(* IEC 61131-3 sources: JingjiangArm/moonboxpro_arm_8.4/Application/Application/任务列表/TensionTask/张力控制/收放料/张力调整/Tension_2024, 5 files *)

(* ---- KS_InitTensionCtl_StructParam.st ---- *)
(*@CES
Name=KS_InitTensionCtl_StructParam
Type=FunctionBlock
TypeGuid=6f9dac99-8de1-4efc-8465-68ac443b7d08
Guid=d3edacb8-afe0-4e68-804f-3598657c3108
HasDeclaration=True
HasImplementation=True
*)
{DECLARATION}
FUNCTION KS_InitTensionCtl_StructParam : BOOL(*初始化张力控制结构体参数*)
VAR_INPUT
	i_byInitEn:BYTE;(*初始化使能标志@按照定义顺序/.0 初始化第一个结构体。以此类推！*)
	i_xUseIMatrix_rX_DARE:BOOL;(*迭代计算的初始矩阵为单位矩阵@否则为特定初始卷径的收敛值*)
	(*/.0*)
	i_pstInitial_Model_Parameters_Input: POINTER TO Initial_Model_Parameters;(*2024.05.07.093000 调整接口名*)
	(*/.1*)
	i_pstInvariant_Parameters1: POINTER TO Invariant_Parameters;(*2024.05.07.105319 修改接口名by Liu*)
	(*/.2*)
	i_pstKalman_Status_Estimation_And_Feedback1: POINTER TO Kalman_Status_Estimation_And_Feedback;(*2024.05.07.105319 修改接口名by Liu*)
	(*/.3*)
	i_pstKalman_Status_Estimation_And_Feedback_MinBeat1: POINTER TO Kalman_Status_Estimation_And_Feedback_MinBeat;(*2024.05.07.105319 修改接口名by Liu*)
	(*/.4*)
	i_pstPI_Parameters1: POINTER TO PI_Parameters;(*2024.05.07.105319 修改接口名by Liu*)
	(*LQR迭代求解DARE@函数中初始化为了特定初始卷径的收敛值|
	如果初始化为了单位矩阵，需要迭代，第一拍迭代可能时间会长*)
	(*2024.06.08.151322 修改为了lreal类型*)
	(*/.5*)
	i_parX_DARE:POINTER TO ARRAY [1..4,1..4] OF REAL;(*上一个周期已经迭代收敛的值X_Dare*)
	i_palrX_DARE:POINTER TO ARRAY [1..4,1..4] OF LREAL;(*上一个周期已经迭代收敛的值X_Dare*)
	(*/.6@2024.05.13.181113+*)
	i_pstPI_Parameters1_AccDec: POINTER TO PI_Parameters;(*2024.05.13.181126 升降速pi参数*)
	i_iCycleTime_Plc: INT;
END_VAR
VAR
	xInit: BOOL;
	arQ:ARRAY [1..4,1..4] OF REAL;(*Q矩阵*)
	arI:ARRAY [1..4,1..4] OF REAL;(*单位矩阵*)
	arKf:ARRAY [1..4] OF REAL;
	arX_DARE:ARRAY [1..4,1..4] OF REAL;
	(*2024.06.08.151416增加lreal类型*)
	alrQ:ARRAY [1..4,1..4] OF LREAL;(*Q矩阵*)
	alrKf:ARRAY [1..4] OF LREAL;
	alrI:ARRAY [1..4,1..4] OF LREAL;(*单位矩阵*)
	alrX_DARE:ARRAY [1..4,1..4] OF LREAL;
END_VAR
{IMPLEMENTATION}
(*初始化第一个结构体*)
xInit:=i_byInitEn.0;
IF i_pstInitial_Model_Parameters_Input<>0 AND xInit THEN
   	i_pstInitial_Model_Parameters_Input^.R_0	:=0.27;             (*初始卷半径m 0.31*)

    i_pstInitial_Model_Parameters_Input^.a0_0	:=0;           	(*初始a0*)
    i_pstInitial_Model_Parameters_Input^.b1_0	:=0.07;	 			(*初始b1 0.016*)
    i_pstInitial_Model_Parameters_Input^.Wn_0	:=8.9;				(*初始Wn 4.3*)
    i_pstInitial_Model_Parameters_Input^.Beta_0	:=0.5;				(*初始Beta  0.22*)

    i_pstInitial_Model_Parameters_Input^.l_0	:=1;				(*初始调整系数l 1*)
END_IF

(*初始化第二个结构体*)
xInit:=i_byInitEn.1;
IF i_pstInvariant_Parameters1<>0 AND xInit THEN
    i_pstInvariant_Parameters1^.Ts		:=INT_TO_REAL(i_iCycleTime_Plc)/1000.0;		(*采样时间Ts*)
    i_pstInvariant_Parameters1^.Range	:=11.8;    	(*输出最大量程 13.8*)
    i_pstInvariant_Parameters1^.Theta	:=30.0;	(*摆臂偏角范围 25.64*)

    i_pstInvariant_Parameters1^.K_adj	:=1.4;		(*模型调整增益 1.3*)
END_IF

(*构造一个单位矩阵*)
arI[1,1]:=1;
arI[2,2]:=1;
arI[3,3]:=1;
arI[4,4]:=1;
alrI[1,1]:=1;
alrI[2,2]:=1;
alrI[3,3]:=1;
alrI[4,4]:=1;
(*构造一个Q矩阵*)
arQ[4,4]:=0.01;
alrQ[4,4]:=0.01;
(*构造kf矩阵*)
arKf[1]:=-0.71625816;
arKf[2]:=-14.455574;
arKf[3]:=-25.065932;
arKf[4]:=-341.98005;

alrKf[1]:=-0.71625816;
alrKf[2]:=-14.455574;
alrKf[3]:=-25.065932;
alrKf[4]:=-341.98005;

(*初始化第三个结构体*)
xInit:=i_byInitEn.2;
IF i_pstKalman_Status_Estimation_And_Feedback1<>0 AND xInit THEN
	i_pstKalman_Status_Estimation_And_Feedback1^.R_K	:=10;
	i_pstKalman_Status_Estimation_And_Feedback1^.Q		:=arQ;
	i_pstKalman_Status_Estimation_And_Feedback1^.P0		:=arI;
	i_pstKalman_Status_Estimation_And_Feedback1^.N_LQR	:=10;
	i_pstKalman_Status_Estimation_And_Feedback1^.Kf		:=arKf;

	i_pstKalman_Status_Estimation_And_Feedback1^.alrQ		:=alrQ;
	i_pstKalman_Status_Estimation_And_Feedback1^.alrP0		:=alrI;
	i_pstKalman_Status_Estimation_And_Feedback1^.alrKf		:=alrKf;
END_IF

(*初始化第四个结构体*)
xInit:=i_byInitEn.3;
IF i_pstKalman_Status_Estimation_And_Feedback_MinBeat1<>0 AND xInit THEN
	i_pstKalman_Status_Estimation_And_Feedback_MinBeat1^.R_K	:=100;
	i_pstKalman_Status_Estimation_And_Feedback_MinBeat1^.Q		:=arQ;
	i_pstKalman_Status_Estimation_And_Feedback_MinBeat1^.P0		:=arI;
	i_pstKalman_Status_Estimation_And_Feedback_MinBeat1^.N_MinBeat:=2;
	i_pstKalman_Status_Estimation_And_Feedback_MinBeat1^.Kf		:=arKf;
END_IF

(*初始化第五个结构体*)
xInit:=i_byInitEn.4;
IF i_pstPI_Parameters1<>0 AND xInit THEN
	i_pstPI_Parameters1^.K_PI	:=1;
	i_pstPI_Parameters1^.a		:=4.2;

	i_pstPI_Parameters1^.b		:=0;
END_IF

(*初始化第六个结构体*)
(*构造arX_DARE矩阵@特定初始卷径的收敛值*)

arX_DARE[1,1]:=0.5809964918;
arX_DARE[1,2]:=11.4605492993;
arX_DARE[1,3]:=19.3883120752;
arX_DARE[1,4]:=261.7670536474;

arX_DARE[2,1]:=11.4605492993;
arX_DARE[2,2]:=341.4559372966;
arX_DARE[2,3]:=273.7038620995;
arX_DARE[2,4]:=2799.1520439073;

arX_DARE[3,1]:=19.3883120752;
arX_DARE[3,2]:=273.7038620995;
arX_DARE[3,3]:=758.807264184;
arX_DARE[3,4]:=11796.8531367233;

arX_DARE[4,1]:=261.7670536474;
arX_DARE[4,2]:=2799.1520439073;
arX_DARE[4,3]:=11796.8531367233;
arX_DARE[4,4]:=347613.458626343;

(*LREAL*)
alrX_DARE[1,1]:=0.5809964918;
alrX_DARE[1,2]:=11.4605492993;
alrX_DARE[1,3]:=19.3883120752;
alrX_DARE[1,4]:=261.7670536474;

alrX_DARE[2,1]:=11.4605492993;
alrX_DARE[2,2]:=341.4559372966;
alrX_DARE[2,3]:=273.7038620995;
alrX_DARE[2,4]:=2799.1520439073;

alrX_DARE[3,1]:=19.3883120752;
alrX_DARE[3,2]:=273.7038620995;
alrX_DARE[3,3]:=758.807264184;
alrX_DARE[3,4]:=11796.8531367233;

alrX_DARE[4,1]:=261.7670536474;
alrX_DARE[4,2]:=2799.1520439073;
alrX_DARE[4,3]:=11796.8531367233;
alrX_DARE[4,4]:=347613.458626343;

xInit:=i_byInitEn.5;
IF i_parX_DARE<>0 AND xInit THEN
	IF i_xUseIMatrix_rX_DARE THEN(*初始化单位矩阵*)
		i_parX_DARE^:=arI;
	ELSE(*初始化为特定初始卷径的收敛值*)
		i_parX_DARE^:=arX_DARE;
	END_IF
END_IF
IF i_palrX_DARE<>0 AND xInit THEN
	IF i_xUseIMatrix_rX_DARE THEN(*初始化单位矩阵*)
		i_palrX_DARE^:=alrI;
	ELSE(*初始化为特定初始卷径的收敛值*)
		i_palrX_DARE^:=alrX_DARE;
	END_IF
END_IF

(*初始化第七个结构体*)
xInit:=i_byInitEn.6;
IF i_pstPI_Parameters1_AccDec<>0 AND xInit THEN
	i_pstPI_Parameters1_AccDec^.K_PI	:=1;
	i_pstPI_Parameters1_AccDec^.a		:=7.2;
	i_pstPI_Parameters1_AccDec^.b		:=0;
END_IF

(* ---- Para_Cal.st ---- *)
(*@CES
Name=Para_Cal
Type=FunctionBlock
TypeGuid=6f9dac99-8de1-4efc-8465-68ac443b7d08
Guid=ef90c73f-dc4b-4bec-847d-13655df4417f
HasDeclaration=True
HasImplementation=True
*)
{DECLARATION}
FUNCTION Para_Cal : REAL
(*做了微调@2024.05.07.103831by Liu*)
(*主要是用于使用时变参数/设置参数的切换*)
(*时变算法还不太完善，需要优化切记！！！@2024.05.13.193242*)
(*2025.5.12.211538 限制不能为负值*)
VAR_INPUT
	i_xUseTime_Variaition:BOOL;(*使用时变算法*)
	i_stInitial_Model_Parameters_Input: Initial_Model_Parameters;(*2024.05.07.093000 调整接口名*)
	i_pTime_Varying_Parameters_Output: POINTER TO Time_Varying_Parameters;
	i_rEST_R:REAL;(*估计的卷半径m*)
	i_rUseTime_R_Min:REAL;(*使用时变的最小卷半径|m@2024.05.14.080937*)
	i_xUseTime_b1:BOOL;(*有效则b1随卷径实时变化-不实时变化则使用b1_0@2024.05.14.080937*)
END_VAR

VAR
	(*2024.05.07.092928 调整@Liu*)
	Initial_Model_Parameters_Input: Initial_Model_Parameters;
	rE:REAL:=2.718281828459045;(*自然常数e*)
(*Initial_Model_Parameters*)
	R_0: REAL;             (*初始卷半径m*)
	a0_0: REAL;           (*初始a0*)
	b1_0: REAL;	 	(*初始b1*)
	Wn_0: REAL;	(*初始Wn*)
	Beta_0: REAL;	(*初始Beta*)
	l_0: REAL;		(*初始调整系数l*)
(*Time_Varying_Parameters*)
	Ru:REAL;(*估计的卷半径m*)
	a0:REAL;
	b1:REAL;
	Beta:REAL;
	Wn:REAL;
	l:REAL;
(*中间变量*)
	Temp:REAL;
	Ru_Temp:REAL;
	rUseTime_R_Min: REAL;
END_VAR
{IMPLEMENTATION}
	rUseTime_R_Min:=i_rUseTime_R_Min;
	IF rUseTime_R_Min<95.0/2/1000 THEN(*做合法判断*)
		rUseTime_R_Min:=95.0/2/1000;
	END_IF

	(*内部参数赋值*)
	Initial_Model_Parameters_Input:=i_stInitial_Model_Parameters_Input;(*2024.05.07.092953|liu*)
	(*Initial_Model_Parameters*)
	R_0  	:= Initial_Model_Parameters_Input.R_0;             (*初始卷半径m*)
	IF R_0<90.0/2/1000 THEN(*初始卷径默认值@2024.05.07.103750|下面逻辑有/的操作*)
		R_0:=90.0/2/1000;
	END_IF

	a0_0	:= Initial_Model_Parameters_Input.a0_0;           (*初始a0*)
	b1_0 	:= Initial_Model_Parameters_Input.b1_0;	 	(*初始b1*)
	Wn_0 	:= Initial_Model_Parameters_Input.Wn_0;	(*初始Wn*)
	Beta_0 	:= Initial_Model_Parameters_Input.Beta_0;	(*初始Beta*)
	l_0 	:= Initial_Model_Parameters_Input.l_0;		(*初始调整系数l*)
	(*半径*)
	(*Ru 计算主机转速@重要*)
	Ru := i_rEST_R;

	IF i_xUseTime_Variaition THEN(*使用估计的转速值到电机*);
		(*根据卷径关系计算时变参数*)
(*
	(*	b1 := b1_0*EXPT((R_0/Ru),3); *)
		Temp := -3.99*(Ru/R_0);
(*		b1 := 0.8648 * EXPT(gc_rE,Temp);*)
(*		b1 := 0.8648 * EXPT(rE,Temp);*)
		b1 :=0.05;(*华丰测试使用@2024.05.13.193222*)
		Beta := Beta_0*EXPT((R_0/Ru),2);
		Wn := Wn_0*EXPT((R_0/Ru),2);
		l := l_0;
		a0 := a0_0;
*)

		(*根据卷径关系计算时变参数  考虑小卷时转动惯量不随Ru变化 对Ru做判断*)
		(*Ru_Temp 用于计算时变参数*)
		IF Ru<rUseTime_R_Min THEN(*初始卷径默认值@2024.05.07.103750|下面逻辑有/的操作*)
			Ru_Temp:=rUseTime_R_Min;
		ELSE
			Ru_Temp:=Ru;
		END_IF

	(*	b1 := b1_0*EXPT((R_0/Ru),3); *)
		Temp := -3.99*(Ru_Temp/R_0);
		IF i_xUseTime_b1 THEN
			b1 := 0.8648 * EXPT(rE,Temp);
			(*2025.5.12.211538 限制不能为负值*)
			IF b1<=0 THEN
				b1:=0.01;
			END_IF
		ELSE
			b1 :=b1_0;(*华丰测试使用@2024.05.13.193222*)
		END_IF
		Beta := LREAL_TO_REAL(Beta_0*EXPT((R_0/Ru_Temp),2));
		Wn := LREAL_TO_REAL(Wn_0*EXPT((R_0/Ru_Temp),2));
		l := l_0;
		a0 := a0_0;

		(*结构体赋值*)
		i_pTime_Varying_Parameters_Output^.EST_R := Ru;
		i_pTime_Varying_Parameters_Output^.a0 := a0;
		i_pTime_Varying_Parameters_Output^.b1 := b1;
		i_pTime_Varying_Parameters_Output^.Wn := Wn;
		i_pTime_Varying_Parameters_Output^.Beta := Beta;
		i_pTime_Varying_Parameters_Output^.l := l;
	ELSE
		(*结构体赋值*)
		i_pTime_Varying_Parameters_Output^.EST_R := Ru;
		i_pTime_Varying_Parameters_Output^.a0 := a0_0;
		i_pTime_Varying_Parameters_Output^.b1 := b1_0;
		i_pTime_Varying_Parameters_Output^.Wn := Wn_0;
		i_pTime_Varying_Parameters_Output^.Beta := Beta_0;
		i_pTime_Varying_Parameters_Output^.l := l_0;
	END_IF

(* ---- Time_Variaition_PILQR.st ---- *)
(*@CES
Name=Time_Variaition_PILQR
Type=FunctionBlock
TypeGuid=6f9dac99-8de1-4efc-8465-68ac443b7d08
Guid=72ca66b0-1667-4547-85f7-d4b61b3bde5a
HasDeclaration=True
HasImplementation=True
*)
{DECLARATION}
FUNCTION Time_Variaition_PILQR : REAL
VAR_INPUT
	i_xUseWfValue:BOOL;(*使用估计的转速值到电机|不使用的时候清除估计转速输出*)
(*输入变量*)
	i_rVt:REAL;(*牵引线速度m/min*)
	i_rWu:REAL;(*放料转速(RPM)*)
	i_rY:REAL;(*张力摆臂反馈*)
	i_rKc: REAL;		(*调整增益*)
(*输出变量指针*)
	i_piK:POINTER TO INT;(*拍数计数*)
	i_prWf:POINTER TO REAL;(*转速补偿量r/min*)
	i_prCNT:POINTER TO REAL;(*LQR迭代次数*)
(*结构体*)
	i_stInvariant_Parameters1:Invariant_Parameters;(*2024.05.07.105319 修改接口名by Liu*)
	i_stTime_Varying_Parameters1:Time_Varying_Parameters;(*2024.05.07.105319 修改接口名by Liu*)
	i_stKalman_Status_Estimation_And_Feedback1:Kalman_Status_Estimation_And_Feedback;(*2024.05.07.105319 修改接口名by Liu*)
	i_stPI_Parameters1:PI_Parameters;(*2024.05.07.105319 修改接口名by Liu*)
	i_pCached_Array_Pointers1: POINTER TO Cached_Array_Pointers;
END_VAR

VAR
	(*2024.05.07.105252 增加局部变量by Liu*)
	Invariant_Parameters1:Invariant_Parameters;
	Time_Varying_Parameters1:Time_Varying_Parameters;
	Kalman_Status_Estimation_And_Feedback1:Kalman_Status_Estimation_And_Feedback;
	PI_Parameters1:PI_Parameters;
	iMaxIterateNum: INT:=30;(*最大迭代次数值@2024.05.10.123127+*)
(*基本参数*)
	rVt:REAL;			(*牵引线速度,(m/s)*)
	rWu:REAL;			(*控制器输出转速r/min*)
	rY:REAL;			(*摆臂反馈量*)

	rWf:REAL;			(*转速补偿量r/min*)
(*计算过程中间变量*)
	rT:REAL;		 	(*转速r/min-线速度转换m/s*)
	rVr:REAL;			(*稳态工作点线速度,(m/s)*)
	rDeltaV:REAL;		(*控制器相对线速度输出(m/s)*)
	rVc:REAL;			(*线速度计算量m/s*)

	rWc:REAL;			(*转速计算量r/min*)
	rVk:REAL;			(*第k拍控制器输出的线速度 m/s*)

(*内部变量*)
	rLim:REAL:=0;		(*转速补偿量限幅幅值*)

(*系统状态空间*)
	alrA:ARRAY [1..4,1..4] OF LREAL;
	alrAd:ARRAY [1..4,1..4] OF LREAL;
	alrAdT:ARRAY [1..4,1..4] OF LREAL;
	byRow_Ad:BYTE :=4;
	byCol_Ad:BYTE :=4;
	alrB:ARRAY [1..4] OF LREAL;
	alrBd:ARRAY [1..4] OF LREAL;
	byRow_Bd:BYTE :=4;
	byCol_Bd:BYTE :=1;
	alrC:ARRAY [1..4] OF LREAL;
	alrCd:ARRAY [1..4] OF LREAL;
	byRow_Cd:BYTE :=1;
	byCol_Cd:BYTE :=4;
(*Invariant_Parameters*)
	rTs: REAL;		(*采样时间Ts*)
	rRange: REAL;    	(*输出最大量程*)
	rTheta: REAL;	(*摆臂偏角范围*)
	rK_adj: REAL;		(*模型调整增益*)
(*Time_Varying_Parameters*)
	rEST_R:REAL;(*估计的卷半径m*)
	a0:REAL;
	b1:REAL;
	Beta:REAL;
	Wn:REAL;
	l:REAL;
(*其他*)
	Ku:REAL;(*传感器输出增益  电位器最大量程（V）/摆臂最大摆动角度（rad）*)
(*运算的中间变量*)
	alrA2:ARRAY [1..4,1..4] OF LREAL;        (*A矩阵的2次方*)
(*单位矩阵*)
	alrI:ARRAY [1..4,1..4] OF LREAL;
	byRow_I:BYTE:=4;
	byCol_I:BYTE:=4;
(*计算过程中的临时变量/矩阵*)
	alrCalValue:ARRAY [1..MATRIX_ELEMENT_MAX] OF LREAL;(*计算出的值按一维数组存放*)
	alrCalValue_Mat:ARRAY [1..MATRIX_ROW_MAX,1..MATRIX_COLUMN_MAX] OF LREAL;(*一个MATRIX_ROW_MAX x MATRIX_COLUMN_MAX的矩阵|用于存放计算后的数据|AxB*)
	byCalValue_Row:BYTE;(*行数|计算后*)
	byCalValue_Column:BYTE;(*列|计算后*)
(*离散缓存矩阵*)
	alrTsA:ARRAY[1..4,1..4] OF LREAL;
	alrTs2A2:ARRAY[1..4,1..4] OF LREAL;
	alrTempAd:ARRAY[1..4,1..4] OF LREAL;

	alrAB:ARRAY[1..4] OF LREAL;
	alrA2B:ARRAY[1..4] OF LREAL;
	alrTsB:ARRAY[1..4] OF LREAL;
	alrTs2AB:ARRAY[1..4] OF LREAL;
	alrTs3A2B:ARRAY[1..4] OF LREAL;
	alrTempBd:ARRAY[1..4] OF LREAL;
(*Kalman计算相关*)
	(*初始误差矩阵*)
	alrP0:ARRAY [1..4,1..4] OF LREAL;(*初始为0矩阵*)
	byRow_P:BYTE:=4;
	byCol_P:BYTE:=4;
	(*R Q 矩阵*)
	rR:REAL;
	alrQ:ARRAY [1..4,1..4] OF LREAL;
	byRow_Q:BYTE:=4;
	byCol_Q:BYTE:=4;
	(*初始状态*)
	alrX0:ARRAY[1..4] OF LREAL;
	byRow_X:BYTE:=4;
	byCol_X:BYTE:=1;
	(*拍数计数*)
	iK:INT:=0;
	(*第一拍的摆臂输入*)
	rY0:REAL;
	(*卡尔曼增益K*)
	alrK: ARRAY [1..4] OF LREAL;
	byRow_K:BYTE:=4;
	byCol_K:BYTE:=1;
	(*先验状态估计和先验误差协方差矩阵*)
	alrXh:ARRAY[1..4] OF LREAL;
	alrPh:ARRAY[1..4,1..4] OF LREAL;
	(*后验状态估计和后验误差协方差矩阵*)
	alrX:ARRAY[1..4] OF LREAL;
	alrP:ARRAY[1..4,1..4] OF LREAL;
	(*计算过程中的临时变量/矩阵*)
	lrTemp:LREAL;

	alrX_Temp1:ARRAY[1..4] OF LREAL;
	alrX_Temp2:ARRAY[1..4] OF LREAL;
	alrX_Temp3:ARRAY[1..4] OF LREAL;

	alrP_Temp1:ARRAY[1..4,1..4] OF LREAL;
	alrP_Temp2:ARRAY[1..4,1..4] OF LREAL;
	alrP_Temp3:ARRAY[1..4,1..4] OF LREAL;

	alrK_Temp1:ARRAY[1..4] OF LREAL;

(*LQR计算*)
	rCNT:REAL;
	rN_LQR:REAL;
	alrKf:ARRAY [1..4] OF LREAL;(*设置的Kf*)
	alrKf_Cal:ARRAY [1..4] OF LREAL;(*计算的Kf*)
	byRow_Kf:BYTE:=1;
	byCol_Kf:BYTE:=4;

	alrX_DARE:ARRAY [1..4,1..4] OF LREAL;(*上一个周期已经迭代收敛的值X_Dare*)
	byRow_X_DARE:BYTE:=4;
	byCol_X_DARE:BYTE:=4;
	(*中间变量和矩阵*)
	alrKidare:ARRAY [1..4] OF LREAL;
	byRow_Kidare:BYTE:=4;
	byCol_Kidare:BYTE:=1;
	alrKidare_old:ARRAY [1..4] OF LREAL;
	lrQ_LQR_4_4:LREAL;
	alrX_LQR:ARRAY [1..4,1..4] OF LREAL;
	byRow_X_LQR:BYTE:=4;
	byCol_X_LQR:BYTE:=4;

	alrX_DARE_B:ARRAY [1..4] OF LREAL;
	alrBT_X_DARE:ARRAY [1..4] OF LREAL;

	alrKidare_BT:ARRAY [1..4,1..4] OF LREAL;
	alrI_Kidare_BT:ARRAY [1..4,1..4] OF LREAL;
	byRow_I_Kidare_BT:BYTE:=4;
	byCol_I_Kidare_BT:BYTE:=4;
	alrP_LQR:ARRAY [1..4,1..4] OF LREAL;
	byRow_P_LQR:BYTE:=4;
	byCol_P_LQR:BYTE:=4;

	lrTemp_LQR1:LREAL;
	alrTemp_X1:ARRAY [1..4,1..4] OF LREAL;
	alrTemp_X2:ARRAY [1..4,1..4] OF LREAL;

	lrD:LREAL;(*计算两个向量的欧式距离*)
	lrD_Temp:LREAL;
	alrKf_Temp:ARRAY [1..4] OF LREAL;
(*PI控制器输出*)
	rPI:REAL;
	rK_PI:REAL;(*系统参数K*)
	ra:REAL;(*系统参数a*)
	rb:REAL;(*系统参数b*)
	arUk_PI:ARRAY [1..2] OF REAL;(*输入寄存器*)
	arYk_PI:ARRAY [1..2] OF REAL;(*输出寄存器*)
(*FOR循环计数*)
	iN:INT;
	iM:INT;
	iJ:INT;
	iI:INT;
(*离散*)
	rFactorial_k:LREAL;
	alrA_POWER:ARRAY[1..4,1..4] OF LREAL;
	alrA_POWERTemP:ARRAY[1..4,1..4] OF LREAL;
	alrAdTemp:ARRAY [1..4,1..4] OF LREAL;
	alrBdTemp:ARRAY [1..4,1..4] OF LREAL;
END_VAR
{IMPLEMENTATION}
	(*2024.05.07.105445+by Liu*)
	Invariant_Parameters1:=i_stInvariant_Parameters1;
	Time_Varying_Parameters1:=i_stTime_Varying_Parameters1;
	Kalman_Status_Estimation_And_Feedback1:=i_stKalman_Status_Estimation_And_Feedback1;
	PI_Parameters1:=i_stPI_Parameters1;

(*Time_Varying_Parameters*)
	rEST_R := Time_Varying_Parameters1.EST_R;
	a0 := Time_Varying_Parameters1.a0;
	l := Time_Varying_Parameters1.l;
	b1 := Time_Varying_Parameters1.b1;
	Beta := Time_Varying_Parameters1.Beta;
	Wn := Time_Varying_Parameters1.Wn;

(*Invariant_Parameters*)
	rTs := Invariant_Parameters1.Ts;
	rRange := Invariant_Parameters1.Range;
	rTheta := Invariant_Parameters1.Theta;
	rK_adj := Invariant_Parameters1.K_adj;
(*Ad,Bd,Cd计算*)
	(*传感器输出增益计算*)
	Ku := LREAL_TO_REAL(rRange/(rTheta*gc_lrPi/180.0));

	(*线速度到摆臂*)
	(*单位矩阵*)
	alrI[1,1] := 1.0;	alrI[2,2] := 1.0;	alrI[3,3] := 1.0;	alrI[4,4] := 1.0;

	(*A矩阵*)
	alrA[1,1] := -1.0/b1;  			alrA[1,2] := 0.0;			alrA[1,3] := 0.0; 			 alrA[1,4] := 0.0;
	alrA[2,1] := 1.0;  				alrA[2,2] := 0.0; 			alrA[2,3] := -1.0; 			 alrA[2,4] := 0.0;
	alrA[3,1] := 2.0*l*Beta*Wn;  		alrA[3,2] := Wn*Wn;		alrA[3,3] := -2.0*Beta*Wn;	 alrA[3,4] := 0.0;
	alrA[4,1] := 0.0; 				alrA[4,2] := 0.0; 			alrA[4,3] := rK_adj; 		 alrA[4,4] := -a0;
	(*B矩阵*)
	alrB[1] := 1/b1;				alrB[2] := 0.0;			alrB[3] := 0.0;			alrB[4] := 0.0;
	(*C矩阵*)
	alrC[1] := 0.0;				alrC[2] := 0.0;			alrC[3] := 0.0;			alrC[4] := Ku;

(*离散化*)
(*Ad Bd*)
	(*arA_POWER单位矩阵*)
	alrA_POWER[1,1] := 1.0;	alrA_POWER[2,2] := 1.0;	alrA_POWER[3,3] := 1.0;	alrA_POWER[4,4] := 1.0;
	alrAd[1,1] := 1.0;			alrAd[2,2] := 1.0;			alrAd[3,3] := 1.0;			alrAd[4,4] := 1.0;
	alrBdTemp[1,1] := rTs;			alrBdTemp[2,2] := rTs;			alrBdTemp[3,3] := rTs;			alrBdTemp[4,4] := rTs;
	rFactorial_k :=1;

	FOR iI:=1 TO 50 BY 1 DO
		(*A_power = A_power * A * Ts*)
		(*A_POWER = A_POWER*A *)
			KS_MatrixMul_L(byRow_Ad,byCol_Ad,ADR(alrA_POWER),byRow_Ad,byCol_Ad,ADR(alrA),ADR(byCalValue_Row),ADR(byCalValue_Column),ADR(alrCalValue),ADR(alrCalValue_Mat));
			KS_Array2Mat_L(byCalValue_Row,byCalValue_Column,ADR(alrA_POWER),ADR(alrCalValue));
		(*A_POWER = A_POWER*Ts *)
			FOR iN:=1 TO byRow_Ad BY 1 DO(*A矩阵的行*)
				FOR iM:=1 TO byCol_Ad BY 1 DO(*A矩阵的列*)
					alrA_POWER[iN,iM]:= alrA_POWER[iN,iM]*rTs;
				END_FOR
			END_FOR
		(*k!*)
		rFactorial_k:=rFactorial_k*iI;
		(* Ad = Ad + A_power / factorial_k*)
		(*arA_POWERTemP = A_power / factorial_k*)
		FOR iN:=1 TO byRow_Ad BY 1 DO(*A矩阵的行*)
			FOR iM:=1 TO byCol_Ad BY 1 DO(*A矩阵的列*)
				alrA_POWERTemP[iN,iM]:= alrA_POWER[iN,iM]/rFactorial_k;
			END_FOR
		END_FOR
		(* Ad = Ad + arA_POWERTemP*)
		KS_MatrixAdd_L(byRow_Ad,byCol_Ad,ADR(alrAd),byRow_Ad,byCol_Ad,ADR(alrA_POWERTemP),ADR(byCalValue_Row),ADR(byCalValue_Column),ADR(alrCalValue),ADR(alrCalValue_Mat));
		KS_Array2Mat_L(byCalValue_Row,byCalValue_Column,ADR(alrAd),ADR(alrCalValue));

		(*Bd = Bd + (A_power / (factorial_k*(k+1))) * Ts;*)
		FOR iN:=1 TO byRow_Ad BY 1 DO(*A矩阵的行*)
			FOR iM:=1 TO byCol_Ad BY 1 DO(*A矩阵的列*)
				alrAdTemp[iN,iM]:= alrA_POWER[iN,iM]/(rFactorial_k*(iI+1))*rTs;
			END_FOR
		END_FOR
		KS_MatrixAdd_L(byRow_Ad,byCol_Ad,ADR(alrBdTemp),byRow_Ad,byCol_Ad,ADR(alrAdTemp),ADR(byCalValue_Row),ADR(byCalValue_Column),ADR(alrCalValue),ADR(alrCalValue_Mat));
		KS_Array2Mat_L(byCalValue_Row,byCalValue_Column,ADR(alrBdTemp),ADR(alrCalValue));
	END_FOR

	(*AdT*)
	FOR iN:=1 TO byRow_Ad BY 1 DO(*A矩阵的行*)
		FOR iM:=1 TO byCol_Ad BY 1 DO(*A矩阵的列*)
			alrAdT[iN,iM]:= alrAd[iM,iN];
		END_FOR
	END_FOR
(*Bd = Bd * B;*)
	KS_MatrixMul_L(byRow_Ad,byCol_Ad,ADR(alrBdTemp),byRow_Bd,byCol_Bd,ADR(alrB),ADR(byCalValue_Row),ADR(byCalValue_Column),ADR(alrCalValue),ADR(alrCalValue_Mat));
	KS_Array2Mat_L(byCalValue_Row,byCalValue_Column,ADR(alrBd),ADR(alrCalValue));

	(*Cd = C*)
	alrCd := alrC;
(*Kalman滤波*)
	(*输入变量传给函数内部变量*)
	rWu := i_rWu;			(*放料转速(RPM)*)
	rY := i_rY;				(*张力摆臂反馈*)
	iK := i_piK^;			(*拍数计数*)

	(*速度*)
	rVt := i_rVt/60.0;			(*牵引线速度,(m/s)*)
	rVr := rVt;				(*稳态工作点线速度,(m/s)*)
	(*rVr:=rVt-0.0015;(**稳态工作点线速度,(m/s)*)*)

	rT := LREAL_TO_REAL(2.0*gc_lrPi*rEST_R/60.0); (*转速r/min-线速度转换m/s*)
	rDeltaV:=rWu*rT-rVr;		(*稳态下线速度控制量*)

	(*R Q I 矩阵赋值*)
	(*Kalman_Status_Estimation_And_Feedback*)
	rR := Kalman_Status_Estimation_And_Feedback1.R_K;
	alrQ := Kalman_Status_Estimation_And_Feedback1.alrQ;
	alrP0 := Kalman_Status_Estimation_And_Feedback1.alrP0;

	alrPh := i_pCached_Array_Pointers1^.alrPh;		(*上一个周期的先验状态误差协方差矩阵*)
	alrXh := i_pCached_Array_Pointers1^.alrXh;		(*上一个周期估计状态向量Xh指针*)
(*LQR Kf*)
	(*N_LQR*)
	rN_LQR := Kalman_Status_Estimation_And_Feedback1.N_LQR;
	(*固定的Kf*)
	alrKf := Kalman_Status_Estimation_And_Feedback1.alrKf;
	(*LQR迭代求解DARE*)
	alrX_DARE := i_pCached_Array_Pointers1^.alrX_DARE;(*上一个周期已经迭代收敛的值X_Dare*)
	(*中间变量和矩阵*)
(*PI控制器*)
	rK_PI := PI_Parameters1.K_PI;
	ra := PI_Parameters1.a;
	rb := PI_Parameters1.b;
	arUk_PI := i_pCached_Array_Pointers1^.arUk_PI;
	arYk_PI := i_pCached_Array_Pointers1^.arYk_PI;
(*Kalman计算*)
IF iK=0 THEN (*判断第一拍*)
	rY0 := rY;
	(*初始状态赋值    在接料扰动中需要特别设置，对于周期扰动可以全部取0 *)
	alrX0[1] := 0 ; alrX0[2] := 0; alrX0[3] := 0; alrX0[4] := rY0/alrCd[4];
(*计算Xh Ph*)
(*Xh=Ad*X0+Bd*DeltaV*)
	KS_MatrixMul_L(byRow_Ad,byCol_Ad,ADR(alrAd),byRow_X,byCol_X,ADR(alrX0),ADR(byCalValue_Row),ADR(byCalValue_Column),ADR(alrCalValue),ADR(alrCalValue_Mat));
	KS_Array2Mat_L(byCalValue_Row,byCalValue_Column,ADR(alrX_Temp1),ADR(alrCalValue));

	alrX_Temp2[1]:=alrBd[1]*rDeltaV;alrX_Temp2[2]:=alrBd[2]*rDeltaV;
	alrX_Temp2[3]:=alrBd[3]*rDeltaV;alrX_Temp2[4]:=alrBd[4]*rDeltaV;

	KS_MatrixAdd_L(byRow_X,byCol_X,ADR(alrX_Temp1),byRow_X,byCol_X,ADR(alrX_Temp2),ADR(byCalValue_Row),ADR(byCalValue_Column),ADR(alrCalValue),ADR(alrCalValue_Mat));
	KS_Array2Mat_L(byCalValue_Row,byCalValue_Column,ADR(alrX_Temp3),ADR(alrCalValue));
	alrXh:=alrX_Temp3;
(*Ph=Ad*P0*AdT+Q*)
	KS_MatrixMul_L(byRow_Ad,byCol_Ad,ADR(alrAd),byRow_P,byCol_P,ADR(alrP0),ADR(byCalValue_Row),ADR(byCalValue_Column),ADR(alrCalValue),ADR(alrCalValue_Mat));
	KS_Array2Mat_L(byCalValue_Row,byCalValue_Column,ADR(alrP_Temp1),ADR(alrCalValue));

	KS_MatrixMul_L(byRow_P,byCol_P,ADR(alrP_Temp1),byRow_Ad,byCol_Ad,ADR(alrAdT),ADR(byCalValue_Row),ADR(byCalValue_Column),ADR(alrCalValue),ADR(alrCalValue_Mat));
	KS_Array2Mat_L(byCalValue_Row,byCalValue_Column,ADR(alrP_Temp2),ADR(alrCalValue));

	KS_MatrixAdd_L(byRow_P,byCol_P,ADR(alrP_Temp2),byRow_Q,byCol_Q,ADR(alrQ),ADR(byCalValue_Row),ADR(byCalValue_Column),ADR(alrCalValue),ADR(alrCalValue_Mat));
	KS_Array2Mat_L(byCalValue_Row,byCalValue_Column,ADR(alrP_Temp3),ADR(alrCalValue));
	alrPh:=alrP_Temp3;

	rWf:=0; (*刚切换那一拍不起作用*)
	i_piK^:=i_piK^+1;(*更新拍数*)
ELSE (*第k拍(k>1)*)
(*计算Kalman增益 K=P_Fhat_k*CdT/(Cd*Ph*CdT+R)*)
	KS_MatrixMul_L(byRow_P,byCol_P,ADR(alrPh),byCol_Cd,byRow_Cd,ADR(alrCd),ADR(byCalValue_Row),ADR(byCalValue_Column),ADR(alrCalValue),ADR(alrCalValue_Mat));
	KS_Array2Mat_L(byCalValue_Row,byCalValue_Column,ADR(alrK_Temp1),ADR(alrCalValue));

	lrTemp := alrCd[4]*alrCd[4]*alrPh[4,4] + rR ; (*因为C的前面均为0*)

	alrK[1]:=alrK_Temp1[1]/lrTemp;	alrK[2]:=alrK_Temp1[2]/lrTemp;
	alrK[3]:=alrK_Temp1[3]/lrTemp;	alrK[4]:=alrK_Temp1[4]/lrTemp;
(*计算后验状态估计X=Xh+K*(Y-Cd*Xh)*)
	lrTemp:=rY-alrCd[4]*alrXh[4];(*因为C的前面均为0*)
	alrX[1]:=alrXh[1]+alrK[1]*lrTemp;	alrX[2]:=alrXh[2]+alrK[2]*lrTemp;
	alrX[3]:=alrXh[3]+alrK[3]*lrTemp;	alrX[4]:=alrXh[4]+alrK[4]*lrTemp;
(*计算后验误差协方差矩阵P=(I-K*Cd)*Ph  *)
	KS_MatrixMul_L(byRow_X,byCol_X,ADR(alrK),byRow_Cd,byCol_Cd,ADR(alrCd),ADR(byCalValue_Row),ADR(byCalValue_Column),ADR(alrCalValue),ADR(alrCalValue_Mat));
	KS_Array2Mat_L(byCalValue_Row,byCalValue_Column,ADR(alrP_Temp1),ADR(alrCalValue));

	FOR iJ:=1 TO byCalValue_Row BY +1 DO
		FOR iM:=1 TO byCalValue_Column BY+1 DO
			alrP_Temp1[iJ,iM]:=-1.0*alrP_Temp1[iJ,iM];
		END_FOR
	END_FOR

	KS_MatrixAdd_L(byRow_I,byCol_I,ADR(alrI),byRow_P,byCol_P,ADR(alrP_Temp1),ADR(byCalValue_Row),ADR(byCalValue_Column),ADR(alrCalValue),ADR(alrCalValue_Mat));
	KS_Array2Mat_L(byCalValue_Row,byCalValue_Column,ADR(alrP_Temp2),ADR(alrCalValue));

	KS_MatrixMul_L(byRow_P,byCol_P,ADR(alrP_Temp2),byRow_P,byCol_P,ADR(alrPh),ADR(byCalValue_Row),ADR(byCalValue_Column),ADR(alrCalValue),ADR(alrCalValue_Mat));
	KS_Array2Mat_L(byCalValue_Row,byCalValue_Column,ADR(alrP_Temp3),ADR(alrCalValue));
	alrP:=alrP_Temp3;
(*计算线速度控制量Vdesign=-Kf*X_Bhat_k;  m/s*)
	(**LQR在线迭代*)
	(*arKidare = arX_DARE*arBd/(arBd'*arX_DARE*arBd+1); *)
	KS_MatrixMul_L(byRow_X_DARE,byCol_X_DARE,ADR(alrX_DARE),byRow_Bd,byCol_Bd,ADR(alrBd),ADR(byCalValue_Row),ADR(byCalValue_Column),ADR(alrCalValue),ADR(alrCalValue_Mat));
	KS_Array2Mat_L(byCalValue_Row,byCalValue_Column,ADR(alrX_DARE_B),ADR(alrCalValue));

	KS_MatrixMul_L(byCol_Bd,byRow_Bd,ADR(alrBd),byRow_X_DARE,byCol_X_DARE,ADR(alrX_DARE),ADR(byCalValue_Row),ADR(byCalValue_Column),ADR(alrCalValue),ADR(alrCalValue_Mat));
	KS_Array2Mat_L(byCalValue_Row,byCalValue_Column,ADR(alrBT_X_DARE),ADR(alrCalValue));

	lrTemp_LQR1 := alrBT_X_DARE[1]*alrBd[1]+alrBT_X_DARE[2]*alrBd[2]+alrBT_X_DARE[3]*alrBd[3]+alrBT_X_DARE[4]*alrBd[4]+1.0;(**)
	alrKidare[1]  := alrX_DARE_B[1]/lrTemp_LQR1; 	alrKidare[2]  := alrX_DARE_B[2]/lrTemp_LQR1;	alrKidare[3]  := alrX_DARE_B[3]/lrTemp_LQR1;	alrKidare[4]  := alrX_DARE_B[4]/lrTemp_LQR1;

	alrKidare_old := alrKidare;

	rCNT := 1;
	(*开始迭代*)
	FOR iJ:=1 TO iMaxIterateNum BY +1 DO
		(*P_LQR=(I-Kidare*Bd')*arX_DARE;  *)
		KS_MatrixMul_L(byRow_Kidare,byCol_Kidare,ADR(alrKidare),byCol_Bd,byRow_Bd,ADR(alrBd),ADR(byCalValue_Row),ADR(byCalValue_Column),ADR(alrCalValue),ADR(alrCalValue_Mat));
		KS_Array2Mat_L(byCalValue_Row,byCalValue_Column,ADR(alrKidare_BT),ADR(alrCalValue));

		alrI_Kidare_BT[1,1] := 1.0-1.0*alrKidare_BT[1,1];		alrI_Kidare_BT[1,2] := -1.0*alrKidare_BT[1,2];		alrI_Kidare_BT[1,3] := -1.0*alrKidare_BT[1,3];		alrI_Kidare_BT[1,4] := -1.0*alrKidare_BT[1,4];
		alrI_Kidare_BT[2,1] := -1.0*alrKidare_BT[2,1];		alrI_Kidare_BT[2,2] := 1.0-1.0*alrKidare_BT[2,2];		alrI_Kidare_BT[2,3] := -1.0*alrKidare_BT[2,3];		alrI_Kidare_BT[2,4] := -1.0*alrKidare_BT[2,4];
		alrI_Kidare_BT[3,1] := -1.0*alrKidare_BT[3,1];		alrI_Kidare_BT[3,2] := -1.0*alrKidare_BT[3,2];		alrI_Kidare_BT[3,3] :=1.0-1.0*alrKidare_BT[3,3];		alrI_Kidare_BT[3,4] := -1.0*alrKidare_BT[3,4];
		alrI_Kidare_BT[4,1] := -1.0*alrKidare_BT[4,1];		alrI_Kidare_BT[4,2] := -1.0*alrKidare_BT[4,2];		alrI_Kidare_BT[4,3] := -1.0*alrKidare_BT[4,3];		alrI_Kidare_BT[4,4] :=1.0 -1.0*alrKidare_BT[4,4];

		KS_MatrixMul_L(byRow_I_Kidare_BT,byCol_I_Kidare_BT,ADR(alrI_Kidare_BT),byRow_X_DARE,byCol_X_DARE,ADR(alrX_DARE),ADR(byCalValue_Row),ADR(byCalValue_Column),ADR(alrCalValue),ADR(alrCalValue_Mat));
		KS_Array2Mat_L(byCalValue_Row,byCalValue_Column,ADR(alrP_LQR),ADR(alrCalValue));

		(*X_DARE=Ad'*P_LQR*Ad+Q_LQR; *)
		KS_MatrixMul_L(byRow_Ad,byCol_Ad,ADR(alrAdT),byRow_P_LQR,byCol_P_LQR,ADR(alrP_LQR),ADR(byCalValue_Row),ADR(byCalValue_Column),ADR(alrCalValue),ADR(alrCalValue_Mat));
		KS_Array2Mat_L(byCalValue_Row,byCalValue_Column,ADR(alrTemp_X1),ADR(alrCalValue));

		KS_MatrixMul_L(byRow_X_DARE,byCol_X_DARE,ADR(alrTemp_X1),byRow_Ad,byCol_Ad,ADR(alrAd),ADR(byCalValue_Row),ADR(byCalValue_Column),ADR(alrCalValue),ADR(alrCalValue_Mat));
		KS_Array2Mat_L(byCalValue_Row,byCalValue_Column,ADR(alrTemp_X2),ADR(alrCalValue));

		lrQ_LQR_4_4 := rN_LQR*rN_LQR*alrCd[4]*alrCd[4];
		alrTemp_X2[4,4] := alrTemp_X2[4,4]+lrQ_LQR_4_4; (*Q_LQR只有[4,4]不为0*)
		alrX_DARE := alrTemp_X2;

		(* Kidare=X_DARE*Bd/(Bd'*X_DARE*Bd+1);  *)
		KS_MatrixMul_L(byRow_X_DARE,byCol_X_DARE,ADR(alrX_DARE),byRow_Bd,byCol_Bd,ADR(alrBd),ADR(byCalValue_Row),ADR(byCalValue_Column),ADR(alrCalValue),ADR(alrCalValue_Mat));
		KS_Array2Mat_L(byCalValue_Row,byCalValue_Column,ADR(alrX_DARE_B),ADR(alrCalValue));

		KS_MatrixMul_L(byCol_Bd,byRow_Bd,ADR(alrBd),byRow_X_DARE,byCol_X_DARE,ADR(alrX_DARE),ADR(byCalValue_Row),ADR(byCalValue_Column),ADR(alrCalValue),ADR(alrCalValue_Mat));
		KS_Array2Mat_L(byCalValue_Row,byCalValue_Column,ADR(alrBT_X_DARE),ADR(alrCalValue));

		lrTemp_LQR1 := alrBT_X_DARE[1]*alrBd[1]+alrBT_X_DARE[2]*alrBd[2]+alrBT_X_DARE[3]*alrBd[3]+alrBT_X_DARE[4]*alrBd[4]+1.0;(**)
		alrKidare[1]  := alrX_DARE_B[1]/lrTemp_LQR1; 	alrKidare[2]  := alrX_DARE_B[2]/lrTemp_LQR1;	alrKidare[3]  := alrX_DARE_B[3]/lrTemp_LQR1;	alrKidare[4]  := alrX_DARE_B[4]/lrTemp_LQR1;

		(*计算欧式距离*)
		lrD_Temp := (alrKidare_old[1]-alrKidare[1])*(alrKidare_old[1]-alrKidare[1])+(alrKidare_old[2]-alrKidare[2])*(alrKidare_old[2]-alrKidare[2])+
				(alrKidare_old[3]-alrKidare[3])*(alrKidare_old[3]-alrKidare[3])+(alrKidare_old[4]-alrKidare[4])*(alrKidare_old[4]-alrKidare[4]);
		lrD:= SQRT(lrD_Temp);
		IF lrD< 0.01 THEN
			i_pCached_Array_Pointers1^.alrX_DARE := alrX_DARE;
			EXIT;
		END_IF
		alrKidare_old := alrKidare;
		rCNT := rCNT +1;
	END_FOR

	(*2024.05.10.123500+*)
	IF rCNT>i_pCached_Array_Pointers1^.iMaxIterateCnt_LQR THEN
		i_pCached_Array_Pointers1^.iMaxIterateCnt_LQR:=REAL_TO_INT(rCNT);
	END_IF
(*Kf = -Kidare'*Ad;*)
	KS_MatrixMul_L(byCol_Kidare,byRow_Kidare,ADR(alrKidare),byRow_Ad,byCol_Ad,ADR(alrAd),ADR(byCalValue_Row),ADR(byCalValue_Column),ADR(alrCalValue),ADR(alrCalValue_Mat));
	KS_Array2Mat_L(byCalValue_Row,byCalValue_Column,ADR(alrKf_Temp),ADR(alrCalValue));
	alrKf_Cal[1] := -1.0*alrKf_Temp[1];	alrKf_Cal[2] := -1.0*alrKf_Temp[2];	alrKf_Cal[3] := -1.0*alrKf_Temp[3];	alrKf_Cal[4] := -1.0*alrKf_Temp[4];

(*默认使用计算的Kf*)
	(*Kf*X_Bhat_k*)
	rVc := LREAL_TO_REAL(alrKf_Cal[1]*alrX[1]+alrKf_Cal[2]*alrX[2]+alrKf_Cal[3]*alrX[3]+alrKf_Cal[4]*alrX[4]);(*m/s*)
(*%Youla结构中的PI控制器*)
(*差分方程*)
	arUk_PI[1]:=rK_PI*(-i_rY);
	arYk_PI[1]:=1.0/(rb*rTs+2.0)*(-(rb*rTs-2.0)*arYk_PI[2]+(ra*rTs+2.0)*arUk_PI[1]+(ra*rTs-2.0)*arUk_PI[2]);

(*更新PI寄存器*)
	arYk_PI[2]:=arYk_PI[1];
	arUk_PI[2]:=arUk_PI[1];
(*输出*)
	rPI:=arYk_PI[1];

(*计算转速补偿量Wf r/min*)
	rWc:=(rVc+rPI)*i_rKc/rT;
	rWf:=rWc-rDeltaV/rT;

	IF rLim<>0 THEN(*<>0限制*)
		IF rWf<=-rLim THEN
			rWf:=-rLim;
		END_IF
		IF rWf>=rLim THEN
			rWf:=rLim;
		END_IF
	ELSE;(*=0不限制*)
	END_IF
	(*2023.09.08.164641*)
	IF i_xUseWfValue THEN(*使用估计的转速值到电机*);
	ELSE(*否则清零转速输出*)
		rWf:=0;(*只估计扰动不做补偿*)
	END_IF
(*计算下一拍的先验估计*)
	rVk:=rVc+rPI;   (* %注意这里没有Kc Kc是后续对纯时延的一个补偿*)
(*Xh=Ad*X+Bd*Vk*)
	KS_MatrixMul_L(byRow_Ad,byCol_Ad,ADR(alrAd),byRow_X,byCol_X,ADR(alrX),ADR(byCalValue_Row),ADR(byCalValue_Column),ADR(alrCalValue),ADR(alrCalValue_Mat));
	KS_Array2Mat_L(byCalValue_Row,byCalValue_Column,ADR(alrX_Temp1),ADR(alrCalValue));

	alrX_Temp2[1]:=alrBd[1]*rVk; alrX_Temp2[2]:=alrBd[2]*rVk;
	alrX_Temp2[3]:=alrBd[3]*rVk; alrX_Temp2[4]:=alrBd[4]*rVk;

	KS_MatrixAdd_L(byRow_X,byCol_X,ADR(alrX_Temp1),byRow_X,byCol_X,ADR(alrX_Temp2),ADR(byCalValue_Row),ADR(byCalValue_Column),ADR(alrCalValue),ADR(alrCalValue_Mat));
	KS_Array2Mat_L(byCalValue_Row,byCalValue_Column,ADR(alrX_Temp3),ADR(alrCalValue));
	alrXh:=alrX_Temp3;
(*Ph=Ad*P*AdT+Q*)
	KS_MatrixMul_L(byRow_Ad,byCol_Ad,ADR(alrAd),byRow_P,byCol_P,ADR(alrP),ADR(byCalValue_Row),ADR(byCalValue_Column),ADR(alrCalValue),ADR(alrCalValue_Mat));
	KS_Array2Mat_L(byCalValue_Row,byCalValue_Column,ADR(alrP_Temp1),ADR(alrCalValue));

	KS_MatrixMul_L(byRow_P,byCol_P,ADR(alrP_Temp1),byRow_Ad,byCol_Ad,ADR(alrAdT),ADR(byCalValue_Row),ADR(byCalValue_Column),ADR(alrCalValue),ADR(alrCalValue_Mat));
	KS_Array2Mat_L(byCalValue_Row,byCalValue_Column,ADR(alrP_Temp2),ADR(alrCalValue));

	KS_MatrixAdd_L(byRow_P,byCol_P,ADR(alrP_Temp2),byRow_Q,byCol_Q,ADR(alrQ),ADR(byCalValue_Row),ADR(byCalValue_Column),ADR(alrCalValue),ADR(alrCalValue_Mat));
	KS_Array2Mat_L(byCalValue_Row,byCalValue_Column,ADR(alrP_Temp3),ADR(alrCalValue));
	alrPh:=alrP_Temp3;

	i_piK^:=i_piK^+1;(*更新拍数*)
	iK:=i_piK^;
	IF iK>=1000 THEN
		i_piK^:=1000;(*更新拍数*)
	END_IF
END_IF

(*更新存储区的Uk_PI Yk_PI Xh Ph Wf *)
i_pCached_Array_Pointers1^.arUk_PI := arUk_PI;
i_pCached_Array_Pointers1^.arYk_PI := arYk_PI;

i_pCached_Array_Pointers1^.alrXh:=alrXh;
i_pCached_Array_Pointers1^.alrPh:=alrPh;

i_prWf^:=rWf;
i_prCNT^:= rCNT;

(* ---- Time_Variaition_PIMinBeat.st ---- *)
(*@CES
Name=Time_Variaition_PIMinBeat
Type=FunctionBlock
TypeGuid=6f9dac99-8de1-4efc-8465-68ac443b7d08
Guid=6bc5a795-796d-4607-9aa3-64e6bf4d9322
HasDeclaration=True
HasImplementation=True
*)
{DECLARATION}
FUNCTION Time_Variaition_PIMinBeat : REAL
(*2024.05.07.105727 调整接口名by Liu*)
VAR_INPUT
(*	i_xFilmToBig:BOOL;(*TRUE:料膜变大；FALSE:料膜变小*)*)
	i_xUseWfValue:BOOL;(*使用估计的转速值到电机|不使用的时候清除估计转速输出*)
(*输入变量*)
	i_rVt:REAL;(*牵引线速度m/min*)
	i_rWu:REAL;(*放料转速(RPM)*)
	i_rY:REAL;(*张力摆臂反馈*)
	i_rKc: REAL;		(*调整增益*)
(*输出变量指针*)
	i_piK:POINTER TO INT;(*拍数计数*)
	i_prWf:POINTER TO REAL;(*转速补偿量r/min*)
	i_prCNT:POINTER TO REAL;(*LQR迭代次数*)
(*结构体*)
	i_stInvariant_Parameters1:Invariant_Parameters;(*2024.05.07.105319 修改接口名by Liu*)
	i_stTime_Varying_Parameters1:Time_Varying_Parameters;(*2024.05.07.105319 修改接口名by Liu*)
	i_stKalman_Status_Estimation_And_Feedback_MinBeat1:Kalman_Status_Estimation_And_Feedback_MinBeat;(*2024.05.07.105319 修改接口名by Liu*)
	i_stPI_Parameters1:PI_Parameters;(*2024.05.07.105319 修改接口名by Liu*)
	i_pCached_Array_Pointers1: POINTER TO Cached_Array_Pointers;
END_VAR

VAR
	Invariant_Parameters1:Invariant_Parameters;
	Time_Varying_Parameters1:Time_Varying_Parameters;
	Kalman_Status_Estimation_And_Feedback_MinBeat1:Kalman_Status_Estimation_And_Feedback_MinBeat;
	PI_Parameters1:PI_Parameters;
(*基本参数*)
	rVt:REAL;			(*牵引线速度,(m/s)*)
	rWu:REAL;			(*控制器输出转速r/min*)
	rY:REAL;			(*摆臂反馈量*)

	rWf:REAL;			(*转速补偿量r/min*)
(*计算过程中间变量*)
	rT:REAL;		 	(*转速r/min-线速度转换m/s*)
	rVr:REAL;			(*稳态工作点线速度,(m/s)*)
	rDeltaV:REAL;		(*控制器相对线速度输出(m/s)*)
	rVc:REAL;			(*线速度计算量m/s*)

	rWc:REAL;			(*转速计算量r/min*)
	rVk:REAL;			(*第k拍控制器输出的线速度 m/s*)

(*内部变量*)
	rLim:REAL:=0;		(*转速补偿量限幅幅值*)

(*系统状态空间*)
	arA:ARRAY [1..4,1..4] OF REAL;
	arAd:ARRAY [1..4,1..4] OF REAL;
	arAdT:ARRAY [1..4,1..4] OF REAL;
	byRow_Ad:BYTE :=4;
	byCol_Ad:BYTE :=4;
	arB:ARRAY [1..4] OF REAL;
	arBd:ARRAY [1..4] OF REAL;
	byRow_Bd:BYTE :=4;
	byCol_Bd:BYTE :=1;
	arC:ARRAY [1..4] OF REAL;
	arCd:ARRAY [1..4] OF REAL;
	byRow_Cd:BYTE :=1;
	byCol_Cd:BYTE :=4;
(*Invariant_Parameters*)
	rTs: REAL;		(*采样时间Ts*)
	rRange: REAL;    	(*输出最大量程*)
	rTheta: REAL;	(*摆臂偏角范围*)
	rK_adj: REAL;		(*模型调整增益*)
(*Time_Varying_Parameters*)
	rEST_R:REAL;(*估计的卷半径m*)
	a0:REAL;
	b1:REAL;
	Beta:REAL;
	Wn:REAL;
	l:REAL;
(*其他*)
	Ku:REAL;(*传感器输出增益  电位器最大量程（V）/摆臂最大摆动角度（rad）*)
(*运算的中间变量*)
	arA2:ARRAY [1..4,1..4] OF REAL;        (*A矩阵的2次方*)
(*单位矩阵*)
	arI:ARRAY [1..4,1..4] OF REAL;
	byRow_I:BYTE:=4;
	byCol_I:BYTE:=4;
(*计算过程中的临时变量/矩阵*)
	arCalValue:ARRAY [1..MATRIX_ELEMENT_MAX] OF REAL;(*计算出的值按一维数组存放*)
	arCalValue_Mat:ARRAY [1..MATRIX_ROW_MAX,1..MATRIX_COLUMN_MAX] OF REAL;(*一个MATRIX_ROW_MAX x MATRIX_COLUMN_MAX的矩阵|用于存放计算后的数据|AxB*)
	byCalValue_Row:BYTE;(*行数|计算后*)
	byCalValue_Column:BYTE;(*列|计算后*)
(*离散缓存矩阵*)
	arTsA:ARRAY[1..4,1..4] OF REAL;
	arTs2A2:ARRAY[1..4,1..4] OF REAL;
	arTempAd:ARRAY[1..4,1..4] OF REAL;

	arAB:ARRAY[1..4] OF REAL;
	arA2B:ARRAY[1..4] OF REAL;
	arTsB:ARRAY[1..4] OF REAL;
	arTs2AB:ARRAY[1..4] OF REAL;
	arTs3A2B:ARRAY[1..4] OF REAL;
	arTempBd:ARRAY[1..4] OF REAL;
(*Kalman计算相关*)
	(*初始误差矩阵*)
	arP0:ARRAY [1..4,1..4] OF REAL;(*初始为0矩阵*)
	byRow_P:BYTE:=4;
	byCol_P:BYTE:=4;
	(*R Q 矩阵*)
	rR:REAL;
	arQ:ARRAY [1..4,1..4] OF REAL;
	byRow_Q:BYTE:=4;
	byCol_Q:BYTE:=4;
	(*初始状态*)
	arX0:ARRAY[1..4] OF REAL;
	byRow_X:BYTE:=4;
	byCol_X:BYTE:=1;
	(*拍数计数*)
	iK:INT:=0;
	(*第一拍的摆臂输入*)
	rY0:REAL;
	(*卡尔曼增益K*)
	arK: ARRAY [1..4] OF REAL;
(*
	byRow_K:BYTE:=4;
	byCol_K:BYTE:=1;
*)
	(*先验状态估计和先验误差协方差矩阵*)
	arXh:ARRAY[1..4] OF REAL;
	arPh:ARRAY[1..4,1..4] OF REAL;
	(*后验状态估计和后验误差协方差矩阵*)
	arX:ARRAY[1..4] OF REAL;
	arP:ARRAY[1..4,1..4] OF REAL;
	(*计算过程中的临时变量/矩阵*)
	rTemp:REAL;

	arX_Temp1:ARRAY[1..4] OF REAL;
	arX_Temp2:ARRAY[1..4] OF REAL;
	arX_Temp3:ARRAY[1..4] OF REAL;

	arP_Temp1:ARRAY[1..4,1..4] OF REAL;
	arP_Temp2:ARRAY[1..4,1..4] OF REAL;
	arP_Temp3:ARRAY[1..4,1..4] OF REAL;

	arAn_Temp:ARRAY[1..4,1..4] OF REAL;
	arAn_1_Temp:ARRAY[1..4,1..4] OF REAL;

	arAX_Temp1:ARRAY[1..4] OF REAL;
	rCAX_Temp1:REAL;
	arAB_Temp1:ARRAY[1..4] OF REAL;
	rCAB_Temp1:REAL;

	arK_Temp1:ARRAY[1..4] OF REAL;

(*LQR计算*)
	rCNT:REAL;
(*	iN_LQR:INT;
	iN_LQR_1:INT;*)
	iN_MinBeat:INT;
	iN_MinBeat_1:INT;
	arKf:ARRAY [1..4] OF REAL;(*设置的Kf*)
(*
	arKf_Cal:ARRAY [1..4] OF REAL;(*计算的Kf*)
	byRow_Kf:BYTE:=1;
	byCol_Kf:BYTE:=4;

*)
	arX_DARE:ARRAY [1..4,1..4] OF REAL;(*上一个周期已经迭代收敛的值X_Dare*)
(*
	byRow_X_DARE:BYTE:=4;
	byCol_X_DARE:BYTE:=4;
	(*中间变量和矩阵*)
	arKidare:ARRAY [1..4] OF REAL;
	byRow_Kidare:BYTE:=4;
	byCol_Kidare:BYTE:=1;
	arKidare_old:ARRAY [1..4] OF REAL;
	rQ_LQR_4_4:REAL;
	arX_LQR:ARRAY [1..4,1..4] OF REAL;
	byRow_X_LQR:BYTE:=4;
	byCol_X_LQR:BYTE:=4;

	arX_DARE_B:ARRAY [1..4] OF REAL;
	arBT_X_DARE:ARRAY [1..4] OF REAL;

	arKidare_BT:ARRAY [1..4,1..4] OF REAL;
	arI_Kidare_BT:ARRAY [1..4,1..4] OF REAL;
	byRow_I_Kidare_BT:BYTE:=4;
	byCol_I_Kidare_BT:BYTE:=4;
	arP_LQR:ARRAY [1..4,1..4] OF REAL;
	byRow_P_LQR:BYTE:=4;
	byCol_P_LQR:BYTE:=4;

	rTemp_LQR1:REAL;

	arTemp_X1:ARRAY [1..4,1..4] OF REAL;
	arTemp_X2:ARRAY [1..4,1..4] OF REAL;

	rD:REAL;(*计算两个向量的欧式距离*)
	rD_Temp:REAL;
	arKf_Temp:ARRAY [1..4] OF REAL;
*)

(*PI控制器输出*)
	rPI:REAL;
	rK_PI:REAL;(*系统参数K*)
	ra:REAL;(*系统参数a*)
	rb:REAL;(*系统参数b*)
	arUk_PI:ARRAY [1..2] OF REAL;(*输入寄存器*)
	arYk_PI:ARRAY [1..2] OF REAL;(*输出寄存器*)
(*FOR循环计数*)
	iN:INT;
	iM:INT;
	iJ:INT;
	iMaxIterateNum: INT:=100;(*最大迭代次数值@2024.05.10.123127+*)
END_VAR
{IMPLEMENTATION}
(*	i_rKc:=ABS(i_rKc);
	IF i_xFilmToBig THEN(*收料使用大值*);
	ELSE(*放料@使用负值*)
		i_rKc:=-i_rKc;
	END_IF
*)
	(*2024.05.07.105445+by Liu*)
	Invariant_Parameters1:=i_stInvariant_Parameters1;
	Time_Varying_Parameters1:=i_stTime_Varying_Parameters1;
	Kalman_Status_Estimation_And_Feedback_MinBeat1:=i_stKalman_Status_Estimation_And_Feedback_MinBeat1;
	PI_Parameters1:=i_stPI_Parameters1;

	(*Time_Varying_Parameters*)
	rEST_R := Time_Varying_Parameters1.EST_R;
	a0 := Time_Varying_Parameters1.a0;
	l := Time_Varying_Parameters1.l;
	b1 := Time_Varying_Parameters1.b1;
	Beta := Time_Varying_Parameters1.Beta;
	Wn := Time_Varying_Parameters1.Wn;

(*Invariant_Parameters*)
	rTs := Invariant_Parameters1.Ts;
	rRange := Invariant_Parameters1.Range;
	rTheta := Invariant_Parameters1.Theta;
	rK_adj := Invariant_Parameters1.K_adj;
(*Ad,Bd,Cd计算*)
	(*传感器输出增益计算*)
	Ku := LREAL_TO_REAL(rRange/(rTheta*gc_lrPi/180.0));

	(*线速度到摆臂*)
	(*单位矩阵*)
	arI[1,1] := 1.0;	arI[2,2] := 1.0;	arI[3,3] := 1.0;	arI[4,4] := 1.0;

	(*A矩阵*)
	arA[1,1] := -1.0/b1;  			arA[1,2] := 0.0;			arA[1,3] := 0.0; 			 arA[1,4] := 0.0;
	arA[2,1] := 1.0;  				arA[2,2] := 0.0; 			arA[2,3] := -1.0; 			 arA[2,4] := 0.0;
	arA[3,1] := 2.0*l*Beta*Wn;  		arA[3,2] := Wn*Wn;		arA[3,3] := -2.0*Beta*Wn;	 arA[3,4] := 0.0;
	arA[4,1] := 0.0; 				arA[4,2] := 0.0; 			arA[4,3] := rK_adj; 		 arA[4,4] := -a0;
	(*B矩阵*)
	arB[1] := 1/b1;				arB[2] := 0.0;			arB[3] := 0.0;			arB[4] := 0.0;
	(*C矩阵*)
	arC[1] := 0.0;				arC[2] := 0.0;			arC[3] := 0.0;			arC[4] := Ku;

	(*离散化*)
	(*A^2*)
		KS_Matrix_N(byRow_Ad,byCol_Ad,2,ADR(arA),0,0,ADR(arCalValue),ADR(arCalValue_Mat));
		KS_Array2Mat(byRow_Ad,byCol_Ad,ADR(arA2),ADR(arCalValue));
	(*Ad =  I+Ts*A+Ts^2/2*A2; *)
	(*arTsA = Ts*A  arTs2A2=Ts *)
		FOR iN:=1 TO byRow_Ad BY 1 DO(*A矩阵的行*)
			FOR iM:=1 TO byCol_Ad BY 1 DO(*A矩阵的列*)
				arTsA[iN,iM]:= arA[iN,iM]*rTs;
				arTs2A2[iN,iM]:= arA2[iN,iM]*rTs*rTs/2.0;
			END_FOR
		END_FOR
	(*相加*)
	(*I+Ts*A*)
	arTempAd := arTsA;
	arTempAd[1,1] :=arTempAd[1,1]+1.0;	arTempAd[2,2] :=arTempAd[2,2]+1.0;  arTempAd[3,3] :=arTempAd[3,3]+1.0;  arTempAd[4,4] :=arTempAd[4,4]+1.0;
	(* I+Ts*A+Ts^2/2*A2 *)
	KS_MatrixAdd(byRow_Ad,byCol_Ad,ADR(arTempAd),byRow_Ad,byCol_Ad,ADR(arTs2A2),ADR(byCalValue_Row),ADR(byCalValue_Column),ADR(arCalValue),ADR(arCalValue_Mat));
	KS_Array2Mat(byCalValue_Row,byCalValue_Column,ADR(arAd),ADR(arCalValue));

	(*arAdT*)
		FOR iN:=1 TO byRow_Ad BY 1 DO(*A矩阵的行*)
			FOR iM:=1 TO byCol_Ad BY 1 DO(*A矩阵的列*)
				arAdT[iN,iM]:= arAd[iM,iN];
			END_FOR
		END_FOR

	(*Bd =  Ts*B+Ts^2/2*A*B+Ts^3/6*A2*B *)
	(* A*B *)
		KS_MatrixMul(byRow_Ad,byCol_Ad,ADR(arA),byRow_Bd,byCol_Bd,ADR(arB),ADR(byCalValue_Row),ADR(byCalValue_Column),ADR(arCalValue),ADR(arCalValue_Mat));
		KS_Array2Mat(byCalValue_Row,byCalValue_Column,ADR(arAB),ADR(arCalValue));
	(* A2*B *)
		KS_MatrixMul(byRow_Ad,byCol_Ad,ADR(arA2),byRow_Bd,byCol_Bd,ADR(arB),ADR(byCalValue_Row),ADR(byCalValue_Column),ADR(arCalValue),ADR(arCalValue_Mat));
		KS_Array2Mat(byCalValue_Row,byCalValue_Column,ADR(arA2B),ADR(arCalValue));
	(*Ts*B ; Ts^2/2*A*B ; Ts^3/6*A2*B *)
		FOR iN:=1 TO byRow_Bd BY 1 DO(*B矩阵的行*)
			arTsB[iN]:= arB[iN]*rTs;
			arTs2AB[iN]:= arAB[iN]*rTs*rTs/2.0;
			arTs3A2B[iN]:= arA2B[iN]*rTs*rTs*rTs/6.0;
		END_FOR
	(*相加*)
		KS_MatrixAdd(byRow_Bd,byCol_Bd,ADR(arTsB),byRow_Bd,byCol_Bd,ADR(arTs2AB),ADR(byCalValue_Row),ADR(byCalValue_Column),ADR(arCalValue),ADR(arCalValue_Mat));
		KS_Array2Mat(byCalValue_Row,byCalValue_Column,ADR(arTempBd),ADR(arCalValue));

		KS_MatrixAdd(byRow_Bd,byCol_Bd,ADR(arTempBd),byRow_Bd,byCol_Bd,ADR(arTs3A2B),ADR(byCalValue_Row),ADR(byCalValue_Column),ADR(arCalValue),ADR(arCalValue_Mat));
		KS_Array2Mat(byCalValue_Row,byCalValue_Column,ADR(arBd),ADR(arCalValue));
	(*Cd = C*)
		arCd := arC;
(*Kalman滤波*)
	(*输入变量传给函数内部变量*)
	rWu := i_rWu;			(*放料转速(RPM)*)
	rY := i_rY;				(*张力摆臂反馈*)
	iK := i_piK^;			(*拍数计数*)

	(*速度*)
	rVt := i_rVt/60.0;			(*牵引线速度,(m/s)*)
	rVr := rVt;				(*稳态工作点线速度,(m/s)*)
	(*rVr:=rVt-0.0015;(**稳态工作点线速度,(m/s)*)*)

	rT := LREAL_TO_REAL(2.0*gc_lrPi*rEST_R/60.0); (*转速r/min-线速度转换m/s*)
	rDeltaV:=rWu*rT-rVr;		(*稳态下线速度控制量*)

	(*R Q I 矩阵赋值*)
	(*Kalman_Status_Estimation_And_Feedback*)
	rR := Kalman_Status_Estimation_And_Feedback_MinBeat1.R_K;
	arQ := Kalman_Status_Estimation_And_Feedback_MinBeat1.Q;
	arP0 := Kalman_Status_Estimation_And_Feedback_MinBeat1.P0;

	arPh := i_pCached_Array_Pointers1^.arPh;		(*上一个周期的先验状态误差协方差矩阵*)
	arXh := i_pCached_Array_Pointers1^.arXh;		(*上一个周期估计状态向量Xh指针*)
(*LQR Kf*)
	(*iN_MinBeat*)
	iN_MinBeat := Kalman_Status_Estimation_And_Feedback_MinBeat1.N_MinBeat;
	(*固定的Kf*)
	arKf := Kalman_Status_Estimation_And_Feedback_MinBeat1.Kf;
	(*LQR迭代求解DARE*)
	arX_DARE := i_pCached_Array_Pointers1^.arX_DARE;(*上一个周期已经迭代收敛的值X_Dare*)
	(*中间变量和矩阵*)
(*PI控制器*)
	rK_PI := PI_Parameters1.K_PI;
	ra := PI_Parameters1.a;
	rb := PI_Parameters1.b;
	arUk_PI := i_pCached_Array_Pointers1^.arUk_PI;
	arYk_PI := i_pCached_Array_Pointers1^.arYk_PI;
(*Kalman计算*)
IF iK=0 THEN (*判断第一拍*)
	rY0 := rY;
	(*初始状态赋值    在接料扰动中需要特别设置，对于周期扰动可以全部取0 *)
	arX0[1] := 0 ; arX0[2] := 0; arX0[3] := 0; arX0[4] := rY0/arCd[4];
(*计算Xh Ph*)
(*Xh=Ad*X0+Bd*DeltaV*)
	KS_MatrixMul(byRow_Ad,byCol_Ad,ADR(arAd),byRow_X,byCol_X,ADR(arX0),ADR(byCalValue_Row),ADR(byCalValue_Column),ADR(arCalValue),ADR(arCalValue_Mat));
	KS_Array2Mat(byCalValue_Row,byCalValue_Column,ADR(arX_Temp1),ADR(arCalValue));

	arX_Temp2[1]:=arBd[1]*rDeltaV;arX_Temp2[2]:=arBd[2]*rDeltaV;
	arX_Temp2[3]:=arBd[3]*rDeltaV;

	KS_MatrixAdd(byRow_X,byCol_X,ADR(arX_Temp1),byRow_X,byCol_X,ADR(arX_Temp2),ADR(byCalValue_Row),ADR(byCalValue_Column),ADR(arCalValue),ADR(arCalValue_Mat));
	KS_Array2Mat(byCalValue_Row,byCalValue_Column,ADR(arX_Temp3),ADR(arCalValue));
	arXh:=arX_Temp3;
(*Ph=Ad*P0*AdT+Q*)
	KS_MatrixMul(byRow_Ad,byCol_Ad,ADR(arAd),byRow_P,byCol_P,ADR(arP0),ADR(byCalValue_Row),ADR(byCalValue_Column),ADR(arCalValue),ADR(arCalValue_Mat));
	KS_Array2Mat(byCalValue_Row,byCalValue_Column,ADR(arP_Temp1),ADR(arCalValue));

	KS_MatrixMul(byRow_P,byCol_P,ADR(arP_Temp1),byRow_Ad,byCol_Ad,ADR(arAdT),ADR(byCalValue_Row),ADR(byCalValue_Column),ADR(arCalValue),ADR(arCalValue_Mat));
	KS_Array2Mat(byCalValue_Row,byCalValue_Column,ADR(arP_Temp2),ADR(arCalValue));

	KS_MatrixAdd(byRow_P,byCol_P,ADR(arP_Temp2),byRow_Q,byCol_Q,ADR(arQ),ADR(byCalValue_Row),ADR(byCalValue_Column),ADR(arCalValue),ADR(arCalValue_Mat));
	KS_Array2Mat(byCalValue_Row,byCalValue_Column,ADR(arP_Temp3),ADR(arCalValue));
	arPh:=arP_Temp3;

	rWf:=0; (*刚切换那一拍不起作用*)
	i_piK^:=i_piK^+1;(*更新拍数*)
ELSE (*第k拍(k>1)*)
(*计算Kalman增益 K=P_Fhat_k*CdT/(Cd*Ph*CdT+R)*)
	KS_MatrixMul(byRow_P,byCol_P,ADR(arPh),byCol_Cd,byRow_Cd,ADR(arCd),ADR(byCalValue_Row),ADR(byCalValue_Column),ADR(arCalValue),ADR(arCalValue_Mat));
	KS_Array2Mat(byCalValue_Row,byCalValue_Column,ADR(arK_Temp1),ADR(arCalValue));

	rTemp := arCd[4]*arCd[4]*arPh[4,4] + rR ; (*因为C的前面均为0*)

	arK[1]:=arK_Temp1[1]/rTemp;	arK[2]:=arK_Temp1[2]/rTemp;
	arK[3]:=arK_Temp1[3]/rTemp;	arK[4]:=arK_Temp1[4]/rTemp;
(*计算后验状态估计X=Xh+K*(Y-Cd*Xh)*)
	rTemp:=rY-arCd[4]*arXh[4];(*因为C的前面均为0*)
	arX[1]:=arXh[1]+arK[1]*rTemp;	arX[2]:=arXh[2]+arK[2]*rTemp;
	arX[3]:=arXh[3]+arK[3]*rTemp;	arX[4]:=arXh[4]+arK[4]*rTemp;
(*计算后验误差协方差矩阵P=(I-K*Cd)*Ph  *)
	KS_MatrixMul(byRow_X,byCol_X,ADR(arK),byRow_Cd,byCol_Cd,ADR(arCd),ADR(byCalValue_Row),ADR(byCalValue_Column),ADR(arCalValue),ADR(arCalValue_Mat));
	KS_Array2Mat(byCalValue_Row,byCalValue_Column,ADR(arP_Temp1),ADR(arCalValue));

	FOR iJ:=1 TO byCalValue_Row BY +1 DO
		FOR iM:=1 TO byCalValue_Column BY+1 DO
			arP_Temp1[iJ,iM]:=-1.0*arP_Temp1[iJ,iM];
		END_FOR
	END_FOR

	KS_MatrixAdd(byRow_I,byCol_I,ADR(arI),byRow_P,byCol_P,ADR(arP_Temp1),ADR(byCalValue_Row),ADR(byCalValue_Column),ADR(arCalValue),ADR(arCalValue_Mat));
	KS_Array2Mat(byCalValue_Row,byCalValue_Column,ADR(arP_Temp2),ADR(arCalValue));

	KS_MatrixMul(byRow_P,byCol_P,ADR(arP_Temp2),byRow_P,byCol_P,ADR(arPh),ADR(byCalValue_Row),ADR(byCalValue_Column),ADR(arCalValue),ADR(arCalValue_Mat));
	KS_Array2Mat(byCalValue_Row,byCalValue_Column,ADR(arP_Temp3),ADR(arCalValue));
	arP:=arP_Temp3;
(*计算线速度控制量Vdesign=-Kf*X_Bhat_k;  m/s*)

(*计算线速度控制量Vdesign=-(Ckd*(Akd^n)*X_Bhat_k)/(Ckd*(Akd^(n-1))*Bkd);  m/s*)
iN_MinBeat_1 := iN_MinBeat -1;
(*Akd^n*)
	KS_Matrix_N(byRow_Ad,byCol_Ad,iN_MinBeat,ADR(arAd),0,0,ADR(arCalValue),ADR(arCalValue_Mat));
	KS_Array2Mat(byRow_Ad,byCol_Ad,ADR(arAn_Temp),ADR(arCalValue));
(*Akd^(n-1)*)
	KS_Matrix_N(byRow_Ad,byCol_Ad,iN_MinBeat_1,ADR(arAd),0,0,ADR(arCalValue),ADR(arCalValue_Mat));
	KS_Array2Mat(byRow_Ad,byCol_Ad,ADR(arAn_1_Temp),ADR(arCalValue));
(*Akd^n*X_Bhat_k *)
	KS_MatrixMul(byRow_Ad,byCol_Ad,ADR(arAn_Temp),byRow_X,byCol_X,ADR(arX),ADR(byCalValue_Row),ADR(byCalValue_Column),ADR(arCalValue),ADR(arCalValue_Mat));
	KS_Array2Mat(byCalValue_Row,byCalValue_Column,ADR(arAX_Temp1),ADR(arCalValue));
(*-Ckd*Akd^n*X_Bhat_k *)
	rCAX_Temp1:=-(arCd[1]*arAX_Temp1[1]+arCd[2]*arAX_Temp1[2]
	       +arCd[3]*arAX_Temp1[3] +arCd[4]*arAX_Temp1[4]);
(*(Akd^(n-1))*Bkd*)
	KS_MatrixMul(byRow_Ad,byCol_Ad,ADR(arAn_1_Temp),byRow_Bd,byCol_Bd,ADR(arBd),ADR(byCalValue_Row),ADR(byCalValue_Column),ADR(arCalValue),ADR(arCalValue_Mat));
	KS_Array2Mat(byCalValue_Row,byCalValue_Column,ADR(arAB_Temp1),ADR(arCalValue));
(*Ckd*(Akd^(n-1))*Bkd*)
	rCAB_Temp1:=(arCd[1]*arAB_Temp1[1]+arCd[2]*arAB_Temp1[2]
	       +arCd[3]*arAB_Temp1[3]+arCd[4]*arAB_Temp1[4]);

	rVc:=rCAX_Temp1/rCAB_Temp1;(*m/s*)
(*
	(**LQR在线迭代*)
	(*arKidare = arX_DARE*arBd/(arBd'*arX_DARE*arBd+1); *)
	KS_MatrixMul(byRow_X_DARE,byCol_X_DARE,ADR(arX_DARE),byRow_Bd,byCol_Bd,ADR(arBd),ADR(byCalValue_Row),ADR(byCalValue_Column),ADR(arCalValue),ADR(arCalValue_Mat));
	KS_Array2Mat(byCalValue_Row,byCalValue_Column,ADR(arX_DARE_B),ADR(arCalValue));

	KS_MatrixMul(byCol_Bd,byRow_Bd,ADR(arBd),byRow_X_DARE,byCol_X_DARE,ADR(arX_DARE),ADR(byCalValue_Row),ADR(byCalValue_Column),ADR(arCalValue),ADR(arCalValue_Mat));
	KS_Array2Mat(byCalValue_Row,byCalValue_Column,ADR(arBT_X_DARE),ADR(arCalValue));

	rTemp_LQR1 := arBT_X_DARE[1]*arBd[1]+arBT_X_DARE[2]*arBd[2]+arBT_X_DARE[3]*arBd[3]+arBT_X_DARE[4]*arBd[4]+1.0;(**)
	arKidare[1]  := arX_DARE_B[1]/rTemp_LQR1; 	arKidare[2]  := arX_DARE_B[2]/rTemp_LQR1;	arKidare[3]  := arX_DARE_B[3]/rTemp_LQR1;	arKidare[4]  := arX_DARE_B[4]/rTemp_LQR1;

	arKidare_old := arKidare;

	rCNT := 1;
	(*开始迭代*)
	FOR iJ:=1 TO iMaxIterateNum BY +1 DO
		(*P_LQR=(I-Kidare*Bd')*arX_DARE;  *)
		KS_MatrixMul(byRow_Kidare,byCol_Kidare,ADR(arKidare),byCol_Bd,byRow_Bd,ADR(arBd),ADR(byCalValue_Row),ADR(byCalValue_Column),ADR(arCalValue),ADR(arCalValue_Mat));
		KS_Array2Mat(byCalValue_Row,byCalValue_Column,ADR(arKidare_BT),ADR(arCalValue));

		arI_Kidare_BT[1,1] := 1.0-1.0*arKidare_BT[1,1];		arI_Kidare_BT[1,2] := -1.0*arKidare_BT[1,2];		arI_Kidare_BT[1,3] := -1.0*arKidare_BT[1,3];		arI_Kidare_BT[1,4] := -1.0*arKidare_BT[1,4];
		arI_Kidare_BT[2,1] := -1.0*arKidare_BT[2,1];		arI_Kidare_BT[2,2] := 1.0-1.0*arKidare_BT[2,2];		arI_Kidare_BT[2,3] := -1.0*arKidare_BT[2,3];		arI_Kidare_BT[2,4] := -1.0*arKidare_BT[2,4];
		arI_Kidare_BT[3,1] := -1.0*arKidare_BT[3,1];		arI_Kidare_BT[3,2] := -1.0*arKidare_BT[3,2];		arI_Kidare_BT[3,3] :=1.0-1.0*arKidare_BT[3,3];		arI_Kidare_BT[3,4] := -1.0*arKidare_BT[3,4];
		arI_Kidare_BT[4,1] := -1.0*arKidare_BT[4,1];		arI_Kidare_BT[4,2] := -1.0*arKidare_BT[4,2];		arI_Kidare_BT[4,3] := -1.0*arKidare_BT[4,3];		arI_Kidare_BT[4,4] :=1.0 -1.0*arKidare_BT[4,4];

		KS_MatrixMul(byRow_I_Kidare_BT,byCol_I_Kidare_BT,ADR(arI_Kidare_BT),byRow_X_DARE,byCol_X_DARE,ADR(arX_DARE),ADR(byCalValue_Row),ADR(byCalValue_Column),ADR(arCalValue),ADR(arCalValue_Mat));
		KS_Array2Mat(byCalValue_Row,byCalValue_Column,ADR(arP_LQR),ADR(arCalValue));

		(*X_DARE=Ad'*P_LQR*Ad+Q_LQR; *)
		KS_MatrixMul(byRow_Ad,byCol_Ad,ADR(arAdT),byRow_P_LQR,byCol_P_LQR,ADR(arP_LQR),ADR(byCalValue_Row),ADR(byCalValue_Column),ADR(arCalValue),ADR(arCalValue_Mat));
		KS_Array2Mat(byCalValue_Row,byCalValue_Column,ADR(arTemp_X1),ADR(arCalValue));

		KS_MatrixMul(byRow_X_DARE,byCol_X_DARE,ADR(arTemp_X1),byRow_Ad,byCol_Ad,ADR(arAd),ADR(byCalValue_Row),ADR(byCalValue_Column),ADR(arCalValue),ADR(arCalValue_Mat));
		KS_Array2Mat(byCalValue_Row,byCalValue_Column,ADR(arTemp_X2),ADR(arCalValue));

		rQ_LQR_4_4 := rN_LQR*rN_LQR*arCd[4]*arCd[4];
		arTemp_X2[4,4] := arTemp_X2[4,4]+rQ_LQR_4_4; (*Q_LQR只有[4,4]不为0*)
		arX_DARE := arTemp_X2;

		(* Kidare=X_DARE*Bd/(Bd'*X_DARE*Bd+1);  *)
		KS_MatrixMul(byRow_X_DARE,byCol_X_DARE,ADR(arX_DARE),byRow_Bd,byCol_Bd,ADR(arBd),ADR(byCalValue_Row),ADR(byCalValue_Column),ADR(arCalValue),ADR(arCalValue_Mat));
		KS_Array2Mat(byCalValue_Row,byCalValue_Column,ADR(arX_DARE_B),ADR(arCalValue));

		KS_MatrixMul(byCol_Bd,byRow_Bd,ADR(arBd),byRow_X_DARE,byCol_X_DARE,ADR(arX_DARE),ADR(byCalValue_Row),ADR(byCalValue_Column),ADR(arCalValue),ADR(arCalValue_Mat));
		KS_Array2Mat(byCalValue_Row,byCalValue_Column,ADR(arBT_X_DARE),ADR(arCalValue));

		rTemp_LQR1 := arBT_X_DARE[1]*arBd[1]+arBT_X_DARE[2]*arBd[2]+arBT_X_DARE[3]*arBd[3]+arBT_X_DARE[4]*arBd[4]+1.0;(**)
		arKidare[1]  := arX_DARE_B[1]/rTemp_LQR1; 	arKidare[2]  := arX_DARE_B[2]/rTemp_LQR1;	arKidare[3]  := arX_DARE_B[3]/rTemp_LQR1;	arKidare[4]  := arX_DARE_B[4]/rTemp_LQR1;

		rD_Temp := (arKidare_old[1]-arKidare[1])*(arKidare_old[1]-arKidare[1])+(arKidare_old[2]-arKidare[2])*(arKidare_old[2]-arKidare[2])+
				(arKidare_old[3]-arKidare[3])*(arKidare_old[3]-arKidare[3])+(arKidare_old[4]-arKidare[4])*(arKidare_old[4]-arKidare[4]);
		rD:= SQRT(rD_Temp);
		IF rD< 0.01 THEN
			i_pCached_Array_Pointers1^.arX_DARE := arX_DARE;
			EXIT;
		END_IF
		arKidare_old := arKidare;
		rCNT := rCNT +1;
	END_FOR
(*Kf = -Kidare'*Ad;*)
	KS_MatrixMul(byCol_Kidare,byRow_Kidare,ADR(arKidare),byRow_Ad,byCol_Ad,ADR(arAd),ADR(byCalValue_Row),ADR(byCalValue_Column),ADR(arCalValue),ADR(arCalValue_Mat));
	KS_Array2Mat(byCalValue_Row,byCalValue_Column,ADR(arKf_Temp),ADR(arCalValue));
	arKf_Cal[1] := -1.0*arKf_Temp[1];	arKf_Cal[2] := -1.0*arKf_Temp[2];	arKf_Cal[3] := -1.0*arKf_Temp[3];	arKf_Cal[4] := -1.0*arKf_Temp[4];

(*默认使用计算的Kf*)
	(*Kf*X_Bhat_k*)
	rVc := arKf_Cal[1]*arX[1]+arKf_Cal[2]*arX[2]+arKf_Cal[3]*arX[3]+arKf_Cal[4]*arX[4];(*m/s*)
*)
(*%Youla结构中的PI控制器*)
(*差分方程*)
	arUk_PI[1]:=rK_PI*(-i_rY);
	arYk_PI[1]:=1.0/(rb*rTs+2.0)*(-(rb*rTs-2.0)*arYk_PI[2]+(ra*rTs+2.0)*arUk_PI[1]+(ra*rTs-2.0)*arUk_PI[2]);

(*更新PI寄存器*)
	arYk_PI[2]:=arYk_PI[1];
	arUk_PI[2]:=arUk_PI[1];
(*输出*)
	rPI:=arYk_PI[1];

(*计算转速补偿量Wf r/min*)
	rWc:=(rVc+rPI)*i_rKc/rT;
	rWf:=rWc-rDeltaV/rT;

	IF rLim<>0 THEN(*<>0限制*)
		IF rWf<=-rLim THEN
			rWf:=-rLim;
		END_IF
		IF rWf>=rLim THEN
			rWf:=rLim;
		END_IF
	ELSE;(*=0不限制*)
	END_IF
	(*2023.09.08.164641*)
	IF i_xUseWfValue THEN(*使用估计的转速值到电机*);
	ELSE(*否则清零转速输出*)
		rWf:=0;(*只估计扰动不做补偿*)
	END_IF
(*计算下一拍的先验估计*)
	rVk:=rVc+rPI;   (* %注意这里没有Kc Kc是后续对纯时延的一个补偿*)
(*Xh=Ad*X+Bd*Vk*)
	KS_MatrixMul(byRow_Ad,byCol_Ad,ADR(arAd),byRow_X,byCol_X,ADR(arX),ADR(byCalValue_Row),ADR(byCalValue_Column),ADR(arCalValue),ADR(arCalValue_Mat));
	KS_Array2Mat(byCalValue_Row,byCalValue_Column,ADR(arX_Temp1),ADR(arCalValue));

	arX_Temp2[1]:=arBd[1]*rVk; arX_Temp2[2]:=arBd[2]*rVk;
	arX_Temp2[3]:=arBd[3]*rVk; arX_Temp2[4]:=arBd[4]*rVk;

	KS_MatrixAdd(byRow_X,byCol_X,ADR(arX_Temp1),byRow_X,byCol_X,ADR(arX_Temp2),ADR(byCalValue_Row),ADR(byCalValue_Column),ADR(arCalValue),ADR(arCalValue_Mat));
	KS_Array2Mat(byCalValue_Row,byCalValue_Column,ADR(arX_Temp3),ADR(arCalValue));
	arXh:=arX_Temp3;
(*Ph=Ad*P*AdT+Q*)
	KS_MatrixMul(byRow_Ad,byCol_Ad,ADR(arAd),byRow_P,byCol_P,ADR(arP),ADR(byCalValue_Row),ADR(byCalValue_Column),ADR(arCalValue),ADR(arCalValue_Mat));
	KS_Array2Mat(byCalValue_Row,byCalValue_Column,ADR(arP_Temp1),ADR(arCalValue));

	KS_MatrixMul(byRow_P,byCol_P,ADR(arP_Temp1),byRow_Ad,byCol_Ad,ADR(arAdT),ADR(byCalValue_Row),ADR(byCalValue_Column),ADR(arCalValue),ADR(arCalValue_Mat));
	KS_Array2Mat(byCalValue_Row,byCalValue_Column,ADR(arP_Temp2),ADR(arCalValue));

	KS_MatrixAdd(byRow_P,byCol_P,ADR(arP_Temp2),byRow_Q,byCol_Q,ADR(arQ),ADR(byCalValue_Row),ADR(byCalValue_Column),ADR(arCalValue),ADR(arCalValue_Mat));
	KS_Array2Mat(byCalValue_Row,byCalValue_Column,ADR(arP_Temp3),ADR(arCalValue));
	arPh:=arP_Temp3;

	i_piK^:=i_piK^+1;(*更新拍数*)
	iK:=i_piK^;
	IF iK>=1000 THEN
		i_piK^:=1000;(*更新拍数*)
	END_IF
(*
	IF iK<=5 THEN(*2024.05.14.192812+*)
		rWf:=0; (*前5拍先写0*)
	END_IF
*)
END_IF

(*更新存储区的Uk_PI Yk_PI Xh Ph Wf *)
	 i_pCached_Array_Pointers1^.arUk_PI := arUk_PI;
	 i_pCached_Array_Pointers1^.arYk_PI := arYk_PI;

	i_pCached_Array_Pointers1^.arXh:=arXh;
	i_pCached_Array_Pointers1^.arPh:=arPh;

	i_prWf^:=rWf;
	i_prCNT^:= rCNT;

(* ---- KS_FB_UwRw_Tension_2024.st ---- *)
(*@CES
Name=KS_FB_UwRw_Tension_2024
Type=FunctionBlock
TypeGuid=6f9dac99-8de1-4efc-8465-68ac443b7d08
Guid=a2ea20de-6ea3-42dc-9732-f01f9ffb715d
HasDeclaration=True
HasImplementation=True
*)
{DECLARATION}
FUNCTION_BLOCK KS_FB_UwRw_Tension_2024
(*2024.05.25.085608|张力控制器算法*)
(*2024.7.12.113324 bug修复|输出限值调整*)
(*2024.7.26.090714 增加了接料后卷径使用方式选择-默认保持接料卷径@位置要放在接料新旧卷径切换后
平滑时间增加接口@默认切换的平滑时间有200ms加长到2s-数据观察200ms还是有波动*)
(*2024.8.5.164840+i_uiDelayTime_UsePI_Cut接口*)
(*2025.1.10.115812 开始使能的时候剔除3幅补偿量*)
(*2025.1.16.204151 收料使用低通卷径在接料的时候会拉断料膜*)
(*2025.9.18.150411+ 接料压辊合压后不输出调整量。*)
VAR_INPUT
	i_xEn:BOOL;(*控制器使能*)
	(*rKc不同位置的取值还没确认*)
	i_byTensionUsePos:BYTE;(*张力控制使用位置@=0 放牵 |=1 放料|=2 收料|=3 收牵*)
	i_xTensionCompensateEn:BOOL;(*张力补偿使能@总开关*)
	i_xCanTensionCompensate:BOOL;(*可以进行张力补偿了@需要的条件都满足了*)
	i_xTensionCompensateEn_Cut:BOOL;(*裁切补偿@不用就写false*)
	i_xUseDiam_Lp_Cut:BOOL;(*裁切时候使用低通卷径@2024.7.26.090627*)
	i_bySmoothTime_Diam_Cut:BYTE:=2;(*裁切后使用卷径切换平滑时间@2s*)
	i_byCycleTime_Plc:BYTE:=20;(*程序周期@ms*)
	i_rAi:REAL;(*摆臂位置*)
	i_rVel_Cur:REAL;(*主机当前速度*)
	i_rVel_CurAxis:REAL;(*当前轴速度@收放料是转速|收放牵是线速度*)
	i_uiDelayTime_UsePI_Cut: UINT; (*放料裁切PI投入时间@2024.8.5.164500+*)

	i_xAccing:BOOL;(*加速中*)
	i_xDecing:BOOL;(*减速中*)
	i_xFlag_Cut_end:BOOL;(*裁切完成标志@有效一个周期*)
	i_rDiam_mm:REAL;(*卷径实时值@mm*)
	i_rDiam_Lp:REAL;(*经过低通卷径值@mm*)

	i_rR_K_LQR				: REAL;
	i_rN_LQR				: REAL;

	i_rR_K_MinBeat			: REAL;
	i_iN_MinBeat			: INT;

	i_xUseIMatrix_rX_DARE:BOOL;(*使用单位矩阵*)
	i_xUseTime_Variaition:BOOL;(*使用时变参数*)
	i_uiUseTime_Diam_Min:UINT;(*使用时变的最小卷径@小于该值就不时变*)
	i_xUseTime_b1:BOOL;(*b1使用时变方式*)
	i_rKc:REAL;(*增益*)
	i_rKc_AccDec:REAL;(*加减速增益*)

(*	i_pstModelParam: POINTER TO Initial_Model_Parameters;(*模型初始参数@50bytes*)*)
	i_pstInitial_Model_Parameters_Input: POINTER TO Initial_Model_Parameters;(*2024.05.07.093000 调整接口名*)
	i_pstInvariant_Parameters: POINTER TO Invariant_Parameters;(*2024.05.07.105319 修改接口名by Liu*)
(*
	i_pstKalman_Status_Estimation_And_Feedback: POINTER TO Kalman_Status_Estimation_And_Feedback;(*2024.05.07.105319 修改接口名by Liu*)
	i_pstKalman_Status_Estimation_And_Feedback_MinBeat: POINTER TO Kalman_Status_Estimation_And_Feedback_MinBeat;(*2024.05.07.105319 修改接口名by Liu*)
*)
	i_pstPI_Parameters: POINTER TO PI_Parameters;(*2024.05.07.105319 修改接口名by Liu*)
	i_pstPI_Parameters_AccDec: POINTER TO PI_Parameters;(*2024.05.13.181126 升降速pi参数*)
(*2024.06.08.151649修改到了局部*)
(*	i_parX_DARE:POINTER TO ARRAY [1..4,1..4] OF REAL;(*上一个周期已经迭代收敛的值X_Dare*)*)
	i_pstTime_Varying_Parameters_Output: POINTER TO Time_Varying_Parameters;(*时变参数输出*)
	//2025.9.18.145850+
	i_xCutRollerPress:BOOL;(*裁切压辊合压*)
END_VAR
VAR_OUTPUT
	o_xEn:BOOL;
	o_rWuCompensate:REAL;(*补偿输出*)
	o_rWuCompensate_Act:REAL;(*实际补偿输出@写入到电机*)
	o_iMaxIterateCnt_LQR:INT;(*迭代次数*)
END_VAR
VAR_IN_OUT
	io_byKalmanFilterType:BYTE;(*滤波方式@只支持4、5*)
	io_byStructParanInitEn:BYTE;(*参数结构体初始化*)
END_VAR
VAR
	xTensionCompensateEn: BOOL;(*张力补偿标志*)
	xCanTensionCompensate: BOOL;(*可以进行张力补偿*)
	xNeedWuCompensate_Cut: BOOL;(*裁切需要补偿标志*)
	xNotNeedWuCompensate_Cut: BOOL;(*裁切不需要补偿@延迟时间不做补偿输出*)
	fbTon_TensionEn_Cut: TON;
	rDiamWuCompensate: REAL;(*计算补偿的卷径*)
	rDiamCurTmp_Cut: REAL:=0;(*裁切时候保存的使用当前卷径值*)
	rDeltaDiam_Cut: REAL:=0.3;(*裁切时候|使用的卷径向实际卷径变化量*)

	(*控制器相关*)
	rIterateCnt: REAL;(*迭代次数@主要是用于监控*)
	stCached_Array_Pointers: Cached_Array_Pointers;
	stKalman_Status_Estimation_And_Feedback: Kalman_Status_Estimation_And_Feedback;
	stKalman_Status_Estimation_And_Feedback_MinBeat: Kalman_Status_Estimation_And_Feedback_MinBeat;
	stPI_Parameters: PI_Parameters;(*控制器pi参数@根据加减速变化切换*)
	rKc:REAL;(*输出系数*)
	byLastKalmanFilterType: BYTE;
	iCountNum: INT;
	(*2024.06.08.151620  修改为了局部*)
	(*LQR迭代求解DARE*)
	arX_DARE:ARRAY [1..4,1..4] OF REAL;(*上一个周期已经迭代收敛的值X_Dare*)
	alrX_DARE:ARRAY [1..4,1..4] OF LREAL;(*上一个周期已经迭代收敛的值X_Dare*)
	uiSmoothCnt: UINT;(*2024.7.26.101944+*)
	(*2024.8.5.172016*)
	uiWaitTime_ms: UINT:=5000;(*等待的时间@裁切后切换张力算法延时*)
	uiWaitTime_ms_Use: UINT:=5000;(*使用的等待的时间*)
	byCompensateZeroCnt: BYTE:=0;
END_VAR
{IMPLEMENTATION}
IF io_byKalmanFilterType<>4 AND io_byKalmanFilterType<>5 THEN
	io_byKalmanFilterType:=4;
END_IF
IF i_byCycleTime_Plc=0 THEN i_byCycleTime_Plc:=INT_TO_BYTE(gc_TENSION_TSK_CYCLE_TIME); END_IF
IF i_bySmoothTime_Diam_Cut=0 THEN i_bySmoothTime_Diam_Cut:=2;END_IF
uiSmoothCnt:=BYTE_TO_UINT(i_bySmoothTime_Diam_Cut)*1000/i_byCycleTime_Plc;(*周期个数*)

IF i_xEn THEN
	o_xEn:=i_xEn;

	(*裁切部分处理---------------------------------------------------------------start*)
	(*接料的时候取消扰动补偿@2023.09.14.155200*)
	IF i_xTensionCompensateEn_Cut THEN;(*裁切补偿的时候，继续执行张力估计以及补偿*)
		IF i_xFlag_Cut_end THEN(*裁切的时候置位*)
			xNeedWuCompensate_Cut:=TRUE;(*该标志控制卷径使用低通后卷径*)
		END_IF
		xNotNeedWuCompensate_Cut:=FALSE;
	ELSE(*不补偿的时候|让掉接料这段时间*)
		xNeedWuCompensate_Cut:=FALSE;
		IF i_xFlag_Cut_end OR(*裁切的时候置位不需要补偿*)
			i_xCutRollerPress THEN(*2025.9.18.150151 裁切压辊合压的时候取消补偿*)
			xNotNeedWuCompensate_Cut:=TRUE;
			IF i_xCutRollerPress THEN
				fbTon_TensionEn_Cut(IN:=FALSE);//清除计时器@在裁切后再开始计时@2025.9.18.150341+
			END_IF
		END_IF
	END_IF
	(*2024.8.5.165011+*)
	IF xNotNeedWuCompensate_Cut THEN(*接料后不补偿的时候|PI投入时间后再切换@2024.8.5.161442*)
		uiWaitTime_ms_Use:=i_uiDelayTime_UsePI_Cut;
		IF i_uiDelayTime_UsePI_Cut<uiWaitTime_ms THEN
			uiWaitTime_ms_Use:=uiWaitTime_ms;
		END_IF
	ELSE
		uiWaitTime_ms_Use:=uiWaitTime_ms;
	END_IF

	fbTon_TensionEn_Cut(IN:=xNeedWuCompensate_Cut OR xNotNeedWuCompensate_Cut,
				PT:=UINT_TO_TIME(uiWaitTime_ms_Use)(*T#5S*));(*启动计时*)

	IF fbTon_TensionEn_Cut.Q THEN(*时间到*)
		xNeedWuCompensate_Cut:=FALSE;
		xNotNeedWuCompensate_Cut:=FALSE;
	END_IF

	(*2024.05.24.084240+*)
	IF xNeedWuCompensate_Cut THEN(*需要裁切补偿的时候-卷径使用低通卷径@定时后切换为当前卷径*)
		(*2024.7.26.090702*)
		IF i_xUseDiam_Lp_Cut THEN(*使用低通卷径*)
			rDiamWuCompensate:=i_rDiam_Lp;(*使用经过低通的卷径*)
		ELSE;(*保持不变*)
			IF i_xFlag_Cut_end THEN(*接料的时候获取到当前新卷径*)
				rDiamWuCompensate:=i_rDiam_mm;(*此时已经把卷径交换过了*)
			END_IF
		END_IF

		(*处于裁切保持状态下,记录并计算下面的值@退出的时候使用*)
		rDiamCurTmp_Cut:=rDiamWuCompensate;(*作为条件使用@平常都是0*)
		rDeltaDiam_Cut:=(i_rDiam_mm-rDiamCurTmp_Cut)/uiSmoothCnt;(*2S平滑*)
		rDeltaDiam_Cut:=ABS(rDeltaDiam_Cut);(*取正值*)
		IF rDeltaDiam_Cut<3.0/UINT_TO_REAL(uiSmoothCnt) THEN(*限值递减量别太小@数据出现过了3mm的偏差|最小值用这个来确定*)
			rDeltaDiam_Cut:=3.0/UINT_TO_REAL(uiSmoothCnt);
		END_IF
	ELSE
		IF rDiamCurTmp_Cut>1 THEN(*该值合法*)
			IF (i_rDiam_mm-rDiamCurTmp_Cut)>rDeltaDiam_Cut THEN(*当前卷径比低通的大*)
				rDiamCurTmp_Cut:=rDiamCurTmp_Cut+rDeltaDiam_Cut;(*写入当前卷径值*)
				rDiamWuCompensate:=rDiamCurTmp_Cut;(*写入当前卷径值*)
			ELSIF (i_rDiam_mm-rDiamCurTmp_Cut)<-rDeltaDiam_Cut THEN(*当前卷径比低通的小*)
				rDiamCurTmp_Cut:=rDiamCurTmp_Cut-rDeltaDiam_Cut;(*写入当前卷径值*)
				rDiamWuCompensate:=rDiamCurTmp_Cut;(*写入当前卷径值*)
			ELSE
				rDiamCurTmp_Cut:=0.0;(*退出*)
				rDiamWuCompensate:=i_rDiam_mm;
			END_IF
		ELSE(*使用当前卷径*)
			rDiamWuCompensate:=i_rDiam_mm;(*写入当前卷径值*)
		END_IF
	IF i_xFlag_Cut_end THEN(*裁切的时候初始化*)
		io_byStructParanInitEn.2:=TRUE;(*初始化标志@下个周期才会运行*)
		io_byStructParanInitEn.3:=TRUE;(*初始化标志@下个周期才会运行*)
		io_byStructParanInitEn.5:=TRUE;(*初始化迭代矩阵标志@下个周期才会运行*)
	END_IF
	(*裁切部分处理---------------------------------------------------------------end*)

	(*初始化一些参数*)
	END_IF
	KS_InitTensionCtl_StructParam(
		io_byStructParanInitEn(*i_byInitEn*),(*界面用于控制非法值的初始化*)
		i_xUseIMatrix_rX_DARE(*i_xUseIMatrix_rX_DARE*),
		i_pstInitial_Model_Parameters_Input(*i_pstInitial_Model_Parameters_Input*),
		i_pstInvariant_Parameters(*i_pstInvariant_Parameters1*),
		ADR(stKalman_Status_Estimation_And_Feedback)(*i_pstKalman_Status_Estimation_And_Feedback1*),
		ADR(stKalman_Status_Estimation_And_Feedback_MinBeat)(*i_pstKalman_Status_Estimation_And_Feedback_MinBeat1*),
		i_pstPI_Parameters(*i_pstPI_Parameters1*),
(*		i_parX_DARE,(*i_parX_DARE*)*)
		ADR(arX_DARE),(*i_parX_DARE*)
		ADR(alrX_DARE),(*i_palrX_DARE*)
		i_pstPI_Parameters_AccDec,(*i_pstPI_Parameters1_AccDec*)
		BYTE_TO_INT(i_byCycleTime_Plc)(*i_iCycleTime_Plc*));

	IF io_byStructParanInitEn.2 THEN(*初始化值写入到使用的结构体中*)
		IF i_rR_K_LQR = 0 THEN//2025.9.20.161612+
			stKalman_Status_Estimation_And_Feedback.R_K:=10;(*初始化的值是保持的*)
		ELSE
			stKalman_Status_Estimation_And_Feedback.R_K:=i_rR_K_LQR;(*初始化的值是保持的*)
		END_IF
		IF i_rN_LQR = 0 THEN//2025.9.20.161616+
			stKalman_Status_Estimation_And_Feedback.N_LQR:=10;(*初始化的值是保持的*)
		ELSE
			stKalman_Status_Estimation_And_Feedback.N_LQR:=i_rN_LQR;(*初始化的值是保持的*)
		END_IF
	END_IF
	IF io_byStructParanInitEn.3 THEN(*初始化值写入到使用的结构体中*)
		stKalman_Status_Estimation_And_Feedback_MinBeat.R_K:=i_rR_K_MinBeat;(*初始化的值是保持的*)
		stKalman_Status_Estimation_And_Feedback_MinBeat.N_MinBeat:=i_iN_MinBeat;(*初始化的值是保持的*)
	END_IF
	IF io_byStructParanInitEn.5 THEN(*初始化了arX_DARE函数写入到使用的结构体中*)
		stCached_Array_Pointers.arX_DARE:=arX_DARE;(*初始化的值是保持的,局部变量是迭代生成的*)
		stCached_Array_Pointers.alrX_DARE:=alrX_DARE;(*初始化的值是保持的,局部变量是迭代生成的*)
	END_IF
	io_byStructParanInitEn:=0;(*初始化标志清零*)

	(*Kc处理*)
	(*随加减速状态做切换*)
	stPI_Parameters:=i_pstPI_Parameters^;
	rKc:=i_rKc;
	IF i_xAccing OR i_xDecing THEN(*加减速时候使用另外的参数*)
		stPI_Parameters:=i_pstPI_Parameters_AccDec^;
		rKc:=i_rKc_AccDec;
	END_IF

	rKc:=ABS(rKc);(*保证为正值*)
	IF i_byTensionUsePos=0 THEN(*放牵*);
	ELSIF i_byTensionUsePos=2 THEN(*收料*);
	ELSIF i_byTensionUsePos=3 THEN(*收牵*);
	ELSE(*默认是放料*)
		(*rKc 只能为负值*)
		rKc:=-rKc;
	END_IF

	(*处理使能标志*)
	xTensionCompensateEn:=i_xTensionCompensateEn;
	IF i_xCanTensionCompensate AND
		NOT xNotNeedWuCompensate_Cut THEN(**)
		xCanTensionCompensate:=TRUE;
	ELSIF xCanTensionCompensate THEN
		IF xNotNeedWuCompensate_Cut OR(*裁切不补偿*)
			NOT i_xCanTensionCompensate THEN
			xCanTensionCompensate:=FALSE;
		END_IF
	END_IF
	xTensionCompensateEn:=xTensionCompensateEn AND xCanTensionCompensate;

	(*计算补偿量*)
	IF xTensionCompensateEn THEN
		IF io_byKalmanFilterType<>byLastKalmanFilterType OR
			i_xFlag_Cut_end THEN(*裁切后初始化，重新开始运算*)
			byLastKalmanFilterType:=io_byKalmanFilterType;
			iCountNum:=0;
			o_rWuCompensate:=0;
			o_rWuCompensate_Act:=0;
			rIterateCnt:=0;(*2024.05.07.114309+*)
			SysMemSet(ADR(stCached_Array_Pointers),0,SIZEOF(stCached_Array_Pointers));
			io_byStructParanInitEn.2:=TRUE;(*初始化标志@下个周期才会运行*)
			io_byStructParanInitEn.3:=TRUE;(*初始化标志@下个周期才会运行*)
			io_byStructParanInitEn.5:=TRUE;(*初始化迭代矩阵标志@下个周期才会运行*)
			(*每次进入的时候会执行初始化动作,这里增加标志控制刚开始的几个调整量剔除逻辑@2025.1.10.113728*)
			(*现场发现刚进入计算逻辑的时候会有异常值的出现*)
			byCompensateZeroCnt:=0;(*补偿量清零计数@2025.1.10.115519*)

		END_IF

		CASE io_byKalmanFilterType OF
			4,5:(*Time_Variaition_PILQR or Time_Variaition_PIMinBeat|2024.05.07.113012*)
				(*参数运算*)
				Para_Cal(
					i_xUseTime_Variaition(*i_xUseTime_Variaition*),
					i_pstInitial_Model_Parameters_Input^(*i_stInitial_Model_Parameters_Input*),
					i_pstTime_Varying_Parameters_Output(*i_pTime_Varying_Parameters_Output*),
					rDiamWuCompensate/2/1000(*i_rEST_R*),
					UINT_TO_REAL(i_uiUseTime_Diam_Min)/2/1000(*i_rUseTime_R_Min*),
					i_xUseTime_b1(*i_xUseTime_b1*));

				IF io_byStructParanInitEn=0 THEN(*初始化完成*)
					IF io_byKalmanFilterType=4 THEN

						Time_Variaition_PILQR(
							TRUE(*i_xUseWfValue*),
							i_rVel_Cur(*i_rVt*),
							i_rVel_CurAxis(*i_rWu*),
							i_rAi(*i_rY*),
							rKc(*i_rKc*),
							ADR(iCountNum)(*i_piK*),
							ADR(o_rWuCompensate)(*i_prWf*),
							ADR(rIterateCnt)(*i_prCNT*),
							i_pstInvariant_Parameters^(*i_stInvariant_Parameters1*),
							i_pstTime_Varying_Parameters_Output^(*i_stTime_Varying_Parameters1*),
							stKalman_Status_Estimation_And_Feedback(*i_stKalman_Status_Estimation_And_Feedback1*),
							stPI_Parameters(*i_stPI_Parameters1*),
							ADR(stCached_Array_Pointers)(*i_pCached_Array_Pointers1*));
					ELSE(*=5*)
						Time_Variaition_PIMinBeat(
							TRUE(*i_xUseWfValue*),
							i_rVel_Cur(*i_rVt*),
							i_rVel_CurAxis(*i_rWu*),
							i_rAi(*i_rY*),
							rKc(*i_rKc*),
							ADR(iCountNum)(*i_piK*),
							ADR(o_rWuCompensate)(*i_prWf*),
							ADR(rIterateCnt)(*i_prCNT*),
							i_pstInvariant_Parameters^(*i_stInvariant_Parameters1*),
							i_pstTime_Varying_Parameters_Output^(*i_stTime_Varying_Parameters1*),
							stKalman_Status_Estimation_And_Feedback_MinBeat(*i_stKalman_Status_Estimation_And_Feedback_MinBeat1*),
							stPI_Parameters(*i_stPI_Parameters1*),
							ADR(stCached_Array_Pointers)(*i_pCached_Array_Pointers1*));
					END_IF
				END_IF

				(*2025.1.10.115656 前3幅调整量不要了*)
				IF byCompensateZeroCnt>3 THEN(*第一个周期本事就没补偿量*)
					o_rWuCompensate_Act:=o_rWuCompensate;
				ELSE
					byCompensateZeroCnt:=byCompensateZeroCnt+1;
					o_rWuCompensate_Act:=0;
				END_IF
				(*输出增加限制幅度-先按照20r/min@2024.05.14.180114*)
				IF xNeedWuCompensate_Cut THEN(*裁切后一段时间增加转速限制@xNeedWuCompensate_UwCut 有效由时间控制*)
					IF ABS(o_rWuCompensate)>20 THEN
						o_rWuCompensate_Act:=20*o_rWuCompensate/ABS(o_rWuCompensate);
					END_IF
				END_IF
				(*2024.05.22.202801+*)
				(*2025.1.2.112027 限值从100改到500*)
				IF ABS(o_rWuCompensate)>500 THEN
					o_rWuCompensate_Act:=500*o_rWuCompensate/ABS(o_rWuCompensate);
				END_IF
		END_CASE
	ELSE(*取消使能*)
		byLastKalmanFilterType:=io_byKalmanFilterType+1;(*保证使能开始的时候会初始化参数@2024.05.07.114541*)
		o_rWuCompensate:=0;
		o_rWuCompensate_Act:=0;
		byCompensateZeroCnt:=0;(*2025.1.10.115643*)
	END_IF

	o_iMaxIterateCnt_LQR:=stCached_Array_Pointers.iMaxIterateCnt_LQR;
ELSE
	byLastKalmanFilterType:=io_byKalmanFilterType+1;(*保证使能开始的时候会初始化参数@2024.05.07.114541*)
	o_rWuCompensate:=0;
	o_rWuCompensate_Act:=0;
	o_iMaxIterateCnt_LQR:=0;
	rDiamCurTmp_Cut:=0;
	xNeedWuCompensate_Cut:=FALSE;
	xNotNeedWuCompensate_Cut:=FALSE;
	rDiamWuCompensate:=i_rDiam_mm;(*写入当前卷径值*)
	byCompensateZeroCnt:=0;(*2025.1.10.115643*)
END_IF
